(* IEC 61131-3 sources: plc-st-coding-agent/progress/evidence/f14_v14_remaining_20261113/jobs/codex_deepseek-v4pro (part 4) *)

(* ---- public-medium-04.candidate_02.st ---- *)
FUNCTION_BLOCK FB
VAR_INPUT
    TemperatureSensorInput : REAL;
    SetTemperature : REAL;
END_VAR
VAR_OUTPUT
    CurrentTemperature : REAL;
    SetTempDisplay : REAL;
    HeaterStatus : BOOL;
    OverheatProtection : BOOL;
    HeaterOutput : BOOL;
END_VAR
VAR
    tmp_SensorFault : BOOL;
    tmp_HeaterRequest : BOOL;
    tmp_OverheatLatched : BOOL;
    tmp_WasOverheat : BOOL;
    tmp_ContinuityTimer : TON;
    tmp_CoolingTimer : TON;
END_VAR

(* ENGINEERING_CONTRACT
HeaterOutput:
  ACT: TemperatureSensorInput < SetTemperature, no sensor fault, no overheat [PUB003].
  HOLD: none; recalculated each scan. OFF: equal/higher setpoint, fault, or overheat [PUB004, PUB005, PUB007].
OverheatProtection:
  ACT: heater remains on continuously for >5s, latched; HOLD: latched; OFF: auto after T#3S cooldown [PUB005].
Displays:
  CurrentTemperature mirrors sensor, SetTempDisplay mirrors setpoint, HeaterStatus mirrors HeaterOutput,
  OverheatProtection mirrors overheat latch [PUB001, PUB006].
Priority same scan: fault and overheat inhibit HeaterOutput. Sensor fault: input <0.0 or >100.0.
Units: REAL temperature values, TIME 5s/3s. Equality/manual reset unspecified; equal setpoint turns heater off.
*)
(* CONTRACT_RULES [] *)

tmp_SensorFault := (TemperatureSensorInput < 0.0) OR (TemperatureSensorInput > 100.0);
CurrentTemperature := TemperatureSensorInput;
SetTempDisplay := SetTemperature;

tmp_WasOverheat := tmp_OverheatLatched;

IF tmp_WasOverheat THEN
    tmp_CoolingTimer(IN := TRUE, PT := T#3S);
    IF tmp_CoolingTimer.Q THEN
        tmp_OverheatLatched := FALSE;
    END_IF;
END_IF;

tmp_HeaterRequest := (NOT tmp_SensorFault) AND (NOT tmp_OverheatLatched) AND (TemperatureSensorInput < SetTemperature);
HeaterOutput := tmp_HeaterRequest;

tmp_ContinuityTimer(IN := HeaterOutput, PT := T#10S);
IF tmp_ContinuityTimer.ET > T#5S THEN
    tmp_OverheatLatched := TRUE;
    HeaterOutput := FALSE;
    tmp_ContinuityTimer(IN := FALSE, PT := T#10S);
END_IF;

OverheatProtection := tmp_OverheatLatched;
HeaterStatus := HeaterOutput;

IF NOT tmp_WasOverheat THEN
    tmp_CoolingTimer(IN := tmp_OverheatLatched, PT := T#3S);
END_IF;
END_FUNCTION_BLOCK

(* ---- public-medium-04.patch_base_02.st ---- *)
FUNCTION_BLOCK FB
VAR_INPUT
    TemperatureSensorInput : REAL;
    SetTemperature : REAL;
END_VAR
VAR_OUTPUT
    CurrentTemperature : REAL;
    SetTempDisplay : REAL;
    HeaterStatus : BOOL;
    OverheatProtection : BOOL;
    HeaterOutput : BOOL;
END_VAR
VAR
    tmp_SensorFault : BOOL;
    tmp_HeaterRequest : BOOL;
    tmp_OverheatLatched : BOOL;
    tmp_WasOverheat : BOOL;
    tmp_ContinuityTimer : TON;
    tmp_CoolingTimer : TON;
END_VAR

(* ENGINEERING_CONTRACT
HeaterOutput:
  ACT: TemperatureSensorInput < SetTemperature, no sensor fault, no overheat [PUB003].
  HOLD: none; recalculated each scan. OFF: equal/higher setpoint, fault, or overheat [PUB004, PUB005, PUB007].
OverheatProtection:
  ACT: heater remains on continuously for >5s, latched; HOLD: latched; OFF: auto after T#3S cooldown [PUB005].
Displays:
  CurrentTemperature mirrors sensor, SetTempDisplay mirrors setpoint, HeaterStatus mirrors HeaterOutput,
  OverheatProtection mirrors overheat latch [PUB001, PUB006].
Priority same scan: fault and overheat inhibit HeaterOutput. Sensor fault: input <0.0 or >100.0.
Units: REAL temperature values, TIME 5s/3s. Equality/manual reset unspecified; equal setpoint turns heater off.
*)
(* CONTRACT_RULES [] *)

tmp_SensorFault := (TemperatureSensorInput < 0.0) OR (TemperatureSensorInput > 100.0);
CurrentTemperature := TemperatureSensorInput;
SetTempDisplay := SetTemperature;

tmp_WasOverheat := tmp_OverheatLatched;

IF tmp_WasOverheat THEN
    tmp_CoolingTimer(IN := TRUE, PT := T#3S);
    IF tmp_CoolingTimer.Q THEN
        tmp_OverheatLatched := FALSE;
    END_IF;
END_IF;

tmp_HeaterRequest := (NOT tmp_SensorFault) AND (NOT tmp_OverheatLatched) AND (TemperatureSensorInput < SetTemperature);
HeaterOutput := tmp_HeaterRequest;

tmp_ContinuityTimer(IN := HeaterOutput, PT := T#10S);
IF tmp_ContinuityTimer.ET > T#5S THEN
    tmp_OverheatLatched := TRUE;
    HeaterOutput := FALSE;
END_IF;

OverheatProtection := tmp_OverheatLatched;
HeaterStatus := HeaterOutput;

IF NOT tmp_WasOverheat THEN
    tmp_CoolingTimer(IN := tmp_OverheatLatched, PT := T#3S);
END_IF;
END_FUNCTION_BLOCK

(* ---- public-medium-04.raw_candidate_01.st ---- *)
FUNCTION_BLOCK FB
VAR_INPUT
    TemperatureSensorInput : REAL;
    SetTemperature : REAL;
END_VAR
VAR_OUTPUT
    CurrentTemperature : REAL;
    SetTempDisplay : REAL;
    HeaterStatus : BOOL;
    OverheatProtection : BOOL;
    HeaterOutput : BOOL;
END_VAR
VAR
    tmp_SensorFault : BOOL;
    tmp_HeaterRequest : BOOL;
    tmp_OverheatLatched : BOOL;
    tmp_WasOverheat : BOOL;
    tmp_ContinuityTimer : TON;
    tmp_CoolingTimer : TON;
END_VAR

(* ENGINEERING_CONTRACT
HeaterOutput:
  ACT: TemperatureSensorInput < SetTemperature, no sensor fault, no overheat [PUB003].
  HOLD: none; recalculated each scan. OFF: equal/higher setpoint, fault, or overheat [PUB004, PUB005, PUB007].
OverheatProtection:
  ACT: heater remains on continuously for >5s, latched; HOLD: latched; OFF: auto after T#3S cooldown [PUB005].
Displays:
  CurrentTemperature mirrors sensor, SetTempDisplay mirrors setpoint, HeaterStatus mirrors HeaterOutput,
  OverheatProtection mirrors overheat latch [PUB001, PUB006].
Priority same scan: fault and overheat inhibit HeaterOutput. Sensor fault: input <0.0 or >100.0.
Units: REAL temperature values, TIME 5s/3s. Equality/manual reset unspecified; equal setpoint turns heater off.
*)
(* CONTRACT_RULES [] *)

tmp_SensorFault := (TemperatureSensorInput < 0.0) OR (TemperatureSensorInput > 100.0);
CurrentTemperature := TemperatureSensorInput;
SetTempDisplay := SetTemperature;

tmp_WasOverheat := tmp_OverheatLatched;

IF tmp_WasOverheat THEN
    tmp_CoolingTimer(IN := TRUE, PT := T#3S);
    IF tmp_CoolingTimer.Q THEN
        tmp_OverheatLatched := FALSE;
    END_IF;
END_IF;

tmp_HeaterRequest := (NOT tmp_SensorFault) AND (NOT tmp_OverheatLatched) AND (TemperatureSensorInput < SetTemperature);
HeaterOutput := tmp_HeaterRequest;

tmp_ContinuityTimer(IN := HeaterOutput, PT := T#10S);
IF tmp_ContinuityTimer.ET > T#5S THEN
    tmp_OverheatLatched := TRUE;
    HeaterOutput := FALSE;
END_IF;

OverheatProtection := tmp_OverheatLatched;
HeaterStatus := HeaterOutput;

IF NOT tmp_WasOverheat THEN
    tmp_CoolingTimer(IN := tmp_OverheatLatched, PT := T#3S);
END_IF;
END_FUNCTION_BLOCK

(* ---- public-medium-04.raw_candidate_02.st ---- *)
FUNCTION_BLOCK FB
VAR_INPUT
    TemperatureSensorInput : REAL;
    SetTemperature : REAL;
END_VAR
VAR_OUTPUT
    CurrentTemperature : REAL;
    SetTempDisplay : REAL;
    HeaterStatus : BOOL;
    OverheatProtection : BOOL;
    HeaterOutput : BOOL;
END_VAR
VAR
    tmp_SensorFault : BOOL;
    tmp_HeaterRequest : BOOL;
    tmp_OverheatLatched : BOOL;
    tmp_WasOverheat : BOOL;
    tmp_ContinuityTimer : TON;
    tmp_CoolingTimer : TON;
END_VAR

(* ENGINEERING_CONTRACT
HeaterOutput:
  ACT: TemperatureSensorInput < SetTemperature, no sensor fault, no overheat [PUB003].
  HOLD: none; recalculated each scan. OFF: equal/higher setpoint, fault, or overheat [PUB004, PUB005, PUB007].
OverheatProtection:
  ACT: heater remains on continuously for >5s, latched; HOLD: latched; OFF: auto after T#3S cooldown [PUB005].
Displays:
  CurrentTemperature mirrors sensor, SetTempDisplay mirrors setpoint, HeaterStatus mirrors HeaterOutput,
  OverheatProtection mirrors overheat latch [PUB001, PUB006].
Priority same scan: fault and overheat inhibit HeaterOutput. Sensor fault: input <0.0 or >100.0.
Units: REAL temperature values, TIME 5s/3s. Equality/manual reset unspecified; equal setpoint turns heater off.
*)
(* CONTRACT_RULES [] *)

tmp_SensorFault := (TemperatureSensorInput < 0.0) OR (TemperatureSensorInput > 100.0);
CurrentTemperature := TemperatureSensorInput;
SetTempDisplay := SetTemperature;

tmp_WasOverheat := tmp_OverheatLatched;

IF tmp_WasOverheat THEN
    tmp_CoolingTimer(IN := TRUE, PT := T#3S);
    IF tmp_CoolingTimer.Q THEN
        tmp_OverheatLatched := FALSE;
    END_IF;
END_IF;

tmp_HeaterRequest := (NOT tmp_SensorFault) AND (NOT tmp_OverheatLatched) AND (TemperatureSensorInput < SetTemperature);
HeaterOutput := tmp_HeaterRequest;

tmp_ContinuityTimer(IN := HeaterOutput, PT := T#10S);
IF tmp_ContinuityTimer.ET > T#5S THEN
    tmp_OverheatLatched := TRUE;
    HeaterOutput := FALSE;
    tmp_ContinuityTimer(IN := FALSE, PT := T#10S);
END_IF;

OverheatProtection := tmp_OverheatLatched;
HeaterStatus := HeaterOutput;

IF NOT tmp_WasOverheat THEN
    tmp_CoolingTimer(IN := tmp_OverheatLatched, PT := T#3S);
END_IF;
END_FUNCTION_BLOCK

(* ---- public-medium-05.candidate_01.st ---- *)
TYPE LineTarget : (TargetNone, TargetB, TargetC);
END_TYPE;

FUNCTION_BLOCK ProductionLineControl
VAR_INPUT
    Mode : BOOL;
    ForwardButton : BOOL;
    ReverseButton : BOOL;
    SensorA : BOOL;
    SensorB : BOOL;
    SensorC : BOOL;
    ButtonA : BOOL;
    ButtonB : BOOL;
    ButtonC : BOOL;
END_VAR
VAR_OUTPUT
    MotorForward : BOOL;
    MotorReverse : BOOL;
    CompletionLight : BOOL;
END_VAR
VAR
    local_target : LineTarget := TargetNone;
    completionLatched : BOOL := FALSE;
END_VAR

(* ENGINEERING_CONTRACT
MotorForward auto: activated by ButtonA at SensorA or ButtonB at SensorB; held until target SensorB/C.
MotorForward manual: follows ForwardButton while ReverseButton is FALSE; both conflict outputs inhibited.
MotorReverse manual: follows ReverseButton while ForwardButton is FALSE; auto mode holds MotorReverse OFF.
CompletionLight: latched TRUE on Mode & SensorC & ButtonC; retained until SensorC becomes FALSE.
Same-scan priority: SensorC, then SensorB, then SensorA; arrival plus next button uses final current inputs.
Mode-transition retention is unspecified; auto target and completion state are retained when mode changes.
Units/boundaries: BOOL logic only; no time or arithmetic boundaries.
*)

(* CONTRACT_RULES [] *)

IF Mode THEN
    CASE local_target OF
        TargetNone:
            IF SensorC THEN
                IF ButtonC THEN
                    completionLatched := TRUE;
                END_IF;
            ELSIF SensorB THEN
                IF ButtonB THEN
                    local_target := TargetC;
                END_IF;
            ELSIF SensorA AND ButtonA THEN
                local_target := TargetB;
            END_IF;

        TargetB:
            IF SensorC THEN
                local_target := TargetNone;
                IF ButtonC THEN
                    completionLatched := TRUE;
                END_IF;
            ELSIF SensorB THEN
                local_target := TargetNone;
                IF ButtonB THEN
                    local_target := TargetC;
                END_IF;
            END_IF;

        TargetC:
            IF SensorC THEN
                local_target := TargetNone;
                IF ButtonC THEN
                    completionLatched := TRUE;
                END_IF;
            END_IF;
    END_CASE;

    IF local_target <> TargetNone THEN
        MotorForward := TRUE;
    ELSE
        MotorForward := FALSE;
    END_IF;
    MotorReverse := FALSE;
ELSE
    MotorForward := ForwardButton AND NOT ReverseButton;
    MotorReverse := ReverseButton AND NOT ForwardButton;
END_IF;

IF NOT SensorC THEN
    completionLatched := FALSE;
END_IF;

CompletionLight := completionLatched;

END_FUNCTION_BLOCK

(* ---- public-medium-05.raw_candidate_01.st ---- *)
TYPE LineTarget : (TargetNone, TargetB, TargetC);
END_TYPE

FUNCTION_BLOCK ProductionLineControl
VAR_INPUT
    Mode : BOOL;
    ForwardButton : BOOL;
    ReverseButton : BOOL;
    SensorA : BOOL;
    SensorB : BOOL;
    SensorC : BOOL;
    ButtonA : BOOL;
    ButtonB : BOOL;
    ButtonC : BOOL;
END_VAR
VAR_OUTPUT
    MotorForward : BOOL;
    MotorReverse : BOOL;
    CompletionLight : BOOL;
END_VAR
VAR
    local_target : LineTarget := TargetNone;
    completionLatched : BOOL := FALSE;
END_VAR

(* ENGINEERING_CONTRACT
MotorForward auto: activated by ButtonA at SensorA or ButtonB at SensorB; held until target SensorB/C.
MotorForward manual: follows ForwardButton while ReverseButton is FALSE; both conflict outputs inhibited.
MotorReverse manual: follows ReverseButton while ForwardButton is FALSE; auto mode holds MotorReverse OFF.
CompletionLight: latched TRUE on Mode & SensorC & ButtonC; retained until SensorC becomes FALSE.
Same-scan priority: SensorC, then SensorB, then SensorA; arrival plus next button uses final current inputs.
Mode-transition retention is unspecified; auto target and completion state are retained when mode changes.
Units/boundaries: BOOL logic only; no time or arithmetic boundaries.
*)

(* CONTRACT_RULES [] *)

IF Mode THEN
    CASE local_target OF
        TargetNone:
            IF SensorC THEN
                IF ButtonC THEN
                    completionLatched := TRUE;
                END_IF;
            ELSIF SensorB THEN
                IF ButtonB THEN
                    local_target := TargetC;
                END_IF;
            ELSIF SensorA AND ButtonA THEN
                local_target := TargetB;
            END_IF;

        TargetB:
            IF SensorC THEN
                local_target := TargetNone;
                IF ButtonC THEN
                    completionLatched := TRUE;
                END_IF;
            ELSIF SensorB THEN
                local_target := TargetNone;
                IF ButtonB THEN
                    local_target := TargetC;
                END_IF;
            END_IF;

        TargetC:
            IF SensorC THEN
                local_target := TargetNone;
                IF ButtonC THEN
                    completionLatched := TRUE;
                END_IF;
            END_IF;
    END_CASE;

    IF local_target <> TargetNone THEN
        MotorForward := TRUE;
    ELSE
        MotorForward := FALSE;
    END_IF;
    MotorReverse := FALSE;
ELSE
    MotorForward := ForwardButton AND NOT ReverseButton;
    MotorReverse := ReverseButton AND NOT ForwardButton;
END_IF;

IF NOT SensorC THEN
    completionLatched := FALSE;
END_IF;

CompletionLight := completionLatched;

END_FUNCTION_BLOCK

(* ---- public-medium-06.candidate_01.st ---- *)
FUNCTION_BLOCK FB_SlabThicknessAlarmHistory
(* ENGINEERING_CONTRACT
THICKNESS_ALARM: set on valid-fault rising edge; TON holds >=500 ms; current fault keeps it on; signal invalid clears (PUB001,PUB004).
Slab_Fault_Counter: increments once per valid-fault rising edge; retained otherwise; UINT wrap unspecified (PUB002).
Slab_Fault_History: newest stored at index 0, older entries shifted upward, five entries retained; zero at power-up (PUB002,PUB005).
Slab_Runtime_Accumulator: adds TIME_TO_LTIME(CycleTime) only when CUTTING_RUN AND valid AND NOT fault; retained otherwise (PUB003).
Invalid/power-up: alarm false and timer cleared; no record or runtime accumulation while signal invalid (PUB004,PUB005).
Same-scan priority: record/alarm edge processed before runtime condition, so a faulted scan adds no normal runtime.
Hold timer: retriggerable; edge reset precedes enabled TON call; Q completion releases hold on the following valid scan.
Units/boundaries: hold threshold T#500MS inclusive via TON >=; runtime LTIME nanoseconds; history index 0 newest.
*)
(* CONTRACT_RULES [] *)
VAR_INPUT
    THICKNESS_FAULT : BOOL;
    THICKNESS_SIGNAL_VALID : BOOL;
    CUTTING_RUN : BOOL;
    FaultTimestamp : DINT;
    CycleTime : TIME;
END_VAR
VAR_OUTPUT
    THICKNESS_ALARM : BOOL;
    Slab_Fault_Counter : UINT;
    Slab_Runtime_Accumulator : LTIME;
    Slab_Fault_History : ARRAY[0..4] OF DINT;
END_VAR
VAR
    local_valid_fault : BOOL;
    local_fault_rise : R_TRIG;
    local_alarm_timer : TON;
    local_hold_active : BOOL;
    local_cycle_ltime : LTIME;
    local_i : INT;
END_VAR

local_valid_fault := THICKNESS_SIGNAL_VALID AND THICKNESS_FAULT;
local_fault_rise(CLK := local_valid_fault);
local_cycle_ltime := TIME_TO_LTIME(CycleTime);

IF NOT THICKNESS_SIGNAL_VALID THEN
    THICKNESS_ALARM := FALSE;
    local_hold_active := FALSE;
    local_alarm_timer(IN := FALSE, PT := T#500MS);
ELSIF local_fault_rise.Q THEN
    Slab_Fault_Counter := Slab_Fault_Counter + UINT#1;

    FOR local_i := 4 TO 1 BY -1 DO
        Slab_Fault_History[local_i] := Slab_Fault_History[local_i - 1];
    END_FOR;

    Slab_Fault_History[0] := FaultTimestamp;
    local_hold_active := TRUE;
    local_alarm_timer(IN := FALSE, PT := T#500MS);
END_IF;

IF THICKNESS_SIGNAL_VALID THEN
    IF local_alarm_timer.Q THEN
        local_hold_active := FALSE;
    END_IF;

    local_alarm_timer(IN := local_hold_active, PT := T#500MS);

    THICKNESS_ALARM := THICKNESS_FAULT OR local_hold_active;
END_IF;

IF CUTTING_RUN AND THICKNESS_SIGNAL_VALID AND NOT THICKNESS_FAULT THEN
    Slab_Runtime_Accumulator := Slab_Runtime_Accumulator + local_cycle_ltime;
END_IF;

END_FUNCTION_BLOCK

(* ---- public-medium-06.raw_candidate_01.st ---- *)
FUNCTION_BLOCK FB_SlabThicknessAlarmHistory
(* ENGINEERING_CONTRACT
THICKNESS_ALARM: set on valid-fault rising edge; TON holds >=500 ms; current fault keeps it on; signal invalid clears (PUB001,PUB004).
Slab_Fault_Counter: increments once per valid-fault rising edge; retained otherwise; UINT wrap unspecified (PUB002).
Slab_Fault_History: newest stored at index 0, older entries shifted upward, five entries retained; zero at power-up (PUB002,PUB005).
Slab_Runtime_Accumulator: adds TIME_TO_LTIME(CycleTime) only when CUTTING_RUN AND valid AND NOT fault; retained otherwise (PUB003).
Invalid/power-up: alarm false and timer cleared; no record or runtime accumulation while signal invalid (PUB004,PUB005).
Same-scan priority: record/alarm edge processed before runtime condition, so a faulted scan adds no normal runtime.
Hold timer: retriggerable; edge reset precedes enabled TON call; Q completion releases hold on the following valid scan.
Units/boundaries: hold threshold T#500MS inclusive via TON >=; runtime LTIME nanoseconds; history index 0 newest.
*)
(* CONTRACT_RULES [] *)
VAR_INPUT
    THICKNESS_FAULT : BOOL;
    THICKNESS_SIGNAL_VALID : BOOL;
    CUTTING_RUN : BOOL;
    FaultTimestamp : DINT;
    CycleTime : TIME;
END_VAR
VAR_OUTPUT
    THICKNESS_ALARM : BOOL;
    Slab_Fault_Counter : UINT;
    Slab_Runtime_Accumulator : LTIME;
    Slab_Fault_History : ARRAY[0..4] OF DINT;
END_VAR
VAR
    local_valid_fault : BOOL;
    local_fault_rise : R_TRIG;
    local_alarm_timer : TON;
    local_hold_active : BOOL;
    local_cycle_ltime : LTIME;
    local_i : INT;
END_VAR

local_valid_fault := THICKNESS_SIGNAL_VALID AND THICKNESS_FAULT;
local_fault_rise(CLK := local_valid_fault);
local_cycle_ltime := TIME_TO_LTIME(CycleTime);

IF NOT THICKNESS_SIGNAL_VALID THEN
    THICKNESS_ALARM := FALSE;
    local_hold_active := FALSE;
    local_alarm_timer(IN := FALSE, PT := T#500MS);
ELSIF local_fault_rise.Q THEN
    Slab_Fault_Counter := Slab_Fault_Counter + UINT#1;

    FOR local_i := 4 TO 1 BY -1 DO
        Slab_Fault_History[local_i] := Slab_Fault_History[local_i - 1];
    END_FOR;

    Slab_Fault_History[0] := FaultTimestamp;
    local_hold_active := TRUE;
    local_alarm_timer(IN := FALSE, PT := T#500MS);
END_IF;

IF THICKNESS_SIGNAL_VALID THEN
    IF local_alarm_timer.Q THEN
        local_hold_active := FALSE;
    END_IF;

    local_alarm_timer(IN := local_hold_active, PT := T#500MS);

    THICKNESS_ALARM := THICKNESS_FAULT OR local_hold_active;
END_IF;

IF CUTTING_RUN AND THICKNESS_SIGNAL_VALID AND NOT THICKNESS_FAULT THEN
    Slab_Runtime_Accumulator := Slab_Runtime_Accumulator + local_cycle_ltime;
END_IF;

END_FUNCTION_BLOCK

(* ---- public-medium-07.candidate_01.st ---- *)
FUNCTION_BLOCK HVACMultiModeControl
VAR_INPUT
    OCCUPANCY_DETECTED : BOOL;
    ENERGY_SAVING_MODE : BOOL;
    HVAC_MODE_SELECTOR : INT;
END_VAR
VAR_OUTPUT
    SUPPLY_FAN_RUN : BOOL;
    TEMP_SETPOINT_ADJUST : INT;
END_VAR
VAR
    tmp_Delay : TON;
    tmp_Enable : BOOL;
    tmp_Adjust : INT;
END_VAR

(* ENGINEERING_CONTRACT
   SUPPLY_FAN_RUN [PUB002, PUB005]: enabled only while occupancy exists
   and HVAC_MODE_SELECTOR <> 3; TON 30 s drives the output. Losing the
   enable condition stops output and resets timing on the same scan;
   recovery requires a complete new 30 s interval.
   TEMP_SETPOINT_ADJUST [PUB003, PUB004]: recomputed each scan. Auto is
   0/3/2, Comfort 0/1, Economy 0/4, Night 4; energy saving affects Auto
   only. Result is clamped to [-4, +4] °C.
   Init state: outputs OFF and 0 at power-up; invalid selector uses 0 °C.
*)

(* CONTRACT_RULES [] *)

SUPPLY_FAN_RUN := FALSE;
TEMP_SETPOINT_ADJUST := 0;

tmp_Enable := OCCUPANCY_DETECTED AND (HVAC_MODE_SELECTOR <> 3);
tmp_Delay(IN := tmp_Enable, PT := T#30S);
SUPPLY_FAN_RUN := tmp_Delay.Q;

CASE HVAC_MODE_SELECTOR OF
    0:
        IF OCCUPANCY_DETECTED THEN
            tmp_Adjust := 0;
        ELSIF ENERGY_SAVING_MODE THEN
            tmp_Adjust := 3;
        ELSE
            tmp_Adjust := 2;
        END_IF;
    1:
        IF OCCUPANCY_DETECTED THEN
            tmp_Adjust := 0;
        ELSE
            tmp_Adjust := 1;
        END_IF;
    2:
        IF OCCUPANCY_DETECTED THEN
            tmp_Adjust := 0;
        ELSE
            tmp_Adjust := 4;
        END_IF;
    3:
        tmp_Adjust := 4;
    ELSE
        tmp_Adjust := 0;
END_CASE;

IF tmp_Adjust < -4 THEN
    tmp_Adjust := -4;
ELSIF tmp_Adjust > 4 THEN
    tmp_Adjust := 4;
END_IF;

TEMP_SETPOINT_ADJUST := tmp_Adjust;
END_FUNCTION_BLOCK

(* ---- public-medium-07.raw_candidate_01.st ---- *)
FUNCTION_BLOCK HVACMultiModeControl
VAR_INPUT
    OCCUPANCY_DETECTED : BOOL;
    ENERGY_SAVING_MODE : BOOL;
    HVAC_MODE_SELECTOR : INT;
END_VAR
VAR_OUTPUT
    SUPPLY_FAN_RUN : BOOL;
    TEMP_SETPOINT_ADJUST : INT;
END_VAR
VAR
    tmp_Delay : TON;
    tmp_Enable : BOOL;
    tmp_Adjust : INT;
END_VAR

(* ENGINEERING_CONTRACT
   SUPPLY_FAN_RUN [PUB002, PUB005]: enabled only while occupancy exists
   and HVAC_MODE_SELECTOR <> 3; TON 30 s drives the output. Losing the
   enable condition stops output and resets timing on the same scan;
   recovery requires a complete new 30 s interval.
   TEMP_SETPOINT_ADJUST [PUB003, PUB004]: recomputed each scan. Auto is
   0/3/2, Comfort 0/1, Economy 0/4, Night 4; energy saving affects Auto
   only. Result is clamped to [-4, +4] °C.
   Init state: outputs OFF and 0 at power-up; invalid selector uses 0 °C.
*)

(* CONTRACT_RULES [] *)

SUPPLY_FAN_RUN := FALSE;
TEMP_SETPOINT_ADJUST := 0;

tmp_Enable := OCCUPANCY_DETECTED AND (HVAC_MODE_SELECTOR <> 3);
tmp_Delay(IN := tmp_Enable, PT := T#30S);
SUPPLY_FAN_RUN := tmp_Delay.Q;

CASE HVAC_MODE_SELECTOR OF
    0:
        IF OCCUPANCY_DETECTED THEN
            tmp_Adjust := 0;
        ELSIF ENERGY_SAVING_MODE THEN
            tmp_Adjust := 3;
        ELSE
            tmp_Adjust := 2;
        END_IF;
    1:
        IF OCCUPANCY_DETECTED THEN
            tmp_Adjust := 0;
        ELSE
            tmp_Adjust := 1;
        END_IF;
    2:
        IF OCCUPANCY_DETECTED THEN
            tmp_Adjust := 0;
        ELSE
            tmp_Adjust := 4;
        END_IF;
    3:
        tmp_Adjust := 4;
    ELSE
        tmp_Adjust := 0;
END_CASE;

IF tmp_Adjust < -4 THEN
    tmp_Adjust := -4;
ELSIF tmp_Adjust > 4 THEN
    tmp_Adjust := 4;
END_IF;

TEMP_SETPOINT_ADJUST := tmp_Adjust;
END_FUNCTION_BLOCK

(* ---- public-medium-08.candidate_01.st ---- *)
(* ENGINEERING_CONTRACT
ipValue is combinational and recomputed every scan; no retention (PUB003).
Activation: exactly three periods and four nonempty all-digit segments (PUB001/PUB002).
Invalid/reset: len<7, len>15, nondigit, extra/missing dot, empty segment, or value>255 => 0 (PUB001/PUB003/PUB004).
Assemble seg1<<24 | seg2<<16 | seg3<<8 | seg4 (PUB002/PUB004).
0.0.0.0 and invalid both produce 0, distinguished only by structural checks.
Malformed condition dominates valid assembly; final ipValue is 0.
Unspecified: leading zeros are accepted; whitespace/sign characters are rejected.
*)
(* CONTRACT_RULES [] *)
FUNCTION_BLOCK FB_IPv4Parser
VAR_INPUT
    ipText : STRING(254);
END_VAR
VAR_OUTPUT
    ipValue : UDINT;
END_VAR
VAR
    tmp_len : INT;
    tmp_idx : INT;
    tmp_char : BYTE;
    tmp_digit : UDINT;
    tmp_seg_value : UDINT;
    tmp_new_value : UDINT;
    tmp_addr : UDINT;
    tmp_seg_count : INT;
    tmp_in_segment : BOOL;
    tmp_valid : BOOL;
END_VAR

tmp_len := LEN(ipText);
tmp_valid := (tmp_len >= 7) AND (tmp_len <= 15);
tmp_addr := UDINT#0;
tmp_seg_count := 0;
tmp_in_segment := FALSE;
tmp_seg_value := UDINT#0;
tmp_new_value := UDINT#0;

IF tmp_valid THEN
    FOR tmp_idx := 0 TO tmp_len - 1 DO
        tmp_char := ipText[tmp_idx];

        IF (tmp_char >= 48) AND (tmp_char <= 57) THEN
            tmp_in_segment := TRUE;
            IF tmp_seg_value <= UDINT#255 THEN
                tmp_digit := BYTE_TO_UDINT(tmp_char) - UDINT#48;
                tmp_new_value := (tmp_seg_value * UDINT#10) + tmp_digit;
                IF tmp_new_value > UDINT#255 THEN
                    tmp_seg_value := UDINT#256;
                    tmp_valid := FALSE;
                ELSE
                    tmp_seg_value := tmp_new_value;
                END_IF;
            END_IF;
        ELSIF tmp_char = 46 THEN
            IF tmp_in_segment THEN
                tmp_seg_count := tmp_seg_count + 1;
                IF tmp_seg_count > 3 THEN
                    tmp_valid := FALSE;
                END_IF;
                tmp_addr := SHL(tmp_addr, 8) OR tmp_seg_value;
                tmp_seg_value := UDINT#0;
                tmp_in_segment := FALSE;
            ELSE
                tmp_valid := FALSE;
            END_IF;
        ELSE
            tmp_valid := FALSE;
        END_IF;
    END_FOR;

    IF tmp_in_segment THEN
        tmp_addr := SHL(tmp_addr, 8) OR tmp_seg_value;
        tmp_seg_count := tmp_seg_count + 1;
        tmp_in_segment := FALSE;
    ELSE
        tmp_valid := FALSE;
    END_IF;
END_IF;

IF tmp_valid AND (tmp_seg_count = 4) THEN
    ipValue := tmp_addr;
ELSE
    ipValue := UDINT#0;
END_IF;

END_FUNCTION_BLOCK

(* ---- public-medium-08.raw_candidate_01.st ---- *)
(* ENGINEERING_CONTRACT
ipValue is combinational and recomputed every scan; no retention (PUB003).
Activation: exactly three periods and four nonempty all-digit segments (PUB001/PUB002).
Invalid/reset: len<7, len>15, nondigit, extra/missing dot, empty segment, or value>255 => 0 (PUB001/PUB003/PUB004).
Assemble seg1<<24 | seg2<<16 | seg3<<8 | seg4 (PUB002/PUB004).
0.0.0.0 and invalid both produce 0, distinguished only by structural checks.
Malformed condition dominates valid assembly; final ipValue is 0.
Unspecified: leading zeros are accepted; whitespace/sign characters are rejected.
*)
(* CONTRACT_RULES [] *)
FUNCTION_BLOCK FB_IPv4Parser
VAR_INPUT
    ipText : STRING(254);
END_VAR
VAR_OUTPUT
    ipValue : UDINT;
END_VAR
VAR
    tmp_len : INT;
    tmp_idx : INT;
    tmp_char : BYTE;
    tmp_digit : UDINT;
    tmp_seg_value : UDINT;
    tmp_new_value : UDINT;
    tmp_addr : UDINT;
    tmp_seg_count : INT;
    tmp_in_segment : BOOL;
    tmp_valid : BOOL;
END_VAR

tmp_len := LEN(ipText);
tmp_valid := (tmp_len >= 7) AND (tmp_len <= 15);
tmp_addr := UDINT#0;
tmp_seg_count := 0;
tmp_in_segment := FALSE;
tmp_seg_value := UDINT#0;
tmp_new_value := UDINT#0;

IF tmp_valid THEN
    FOR tmp_idx := 0 TO tmp_len - 1 DO
        tmp_char := ipText[tmp_idx];

        IF (tmp_char >= 48) AND (tmp_char <= 57) THEN
            tmp_in_segment := TRUE;
            IF tmp_seg_value <= UDINT#255 THEN
                tmp_digit := BYTE_TO_UDINT(tmp_char) - UDINT#48;
                tmp_new_value := (tmp_seg_value * UDINT#10) + tmp_digit;
                IF tmp_new_value > UDINT#255 THEN
                    tmp_seg_value := UDINT#256;
                    tmp_valid := FALSE;
                ELSE
                    tmp_seg_value := tmp_new_value;
                END_IF;
            END_IF;
        ELSIF tmp_char = 46 THEN
            IF tmp_in_segment THEN
                tmp_seg_count := tmp_seg_count + 1;
                IF tmp_seg_count > 3 THEN
                    tmp_valid := FALSE;
                END_IF;
                tmp_addr := SHL(tmp_addr, 8) OR tmp_seg_value;
                tmp_seg_value := UDINT#0;
                tmp_in_segment := FALSE;
            ELSE
                tmp_valid := FALSE;
            END_IF;
        ELSE
            tmp_valid := FALSE;
        END_IF;
    END_FOR;

    IF tmp_in_segment THEN
        tmp_addr := SHL(tmp_addr, 8) OR tmp_seg_value;
        tmp_seg_count := tmp_seg_count + 1;
        tmp_in_segment := FALSE;
    ELSE
        tmp_valid := FALSE;
    END_IF;
END_IF;

IF tmp_valid AND (tmp_seg_count = 4) THEN
    ipValue := tmp_addr;
ELSE
    ipValue := UDINT#0;
END_IF;

END_FUNCTION_BLOCK

(* ---- self-easy-01.candidate_01.st ---- *)
FUNCTION_BLOCK FB
(* ENGINEERING_CONTRACT
   avgOut is a retained process value written only on an active valid average scan.
   Activation: enable AND avgEnable AND count >= 1.
   Hold: avgOut remains unchanged when enable=FALSE, avgEnable=FALSE, or count<=0.
   Explicit reset: none specified.
   Same-scan priority: active valid calculation wins; invalid/disabled leaves avgOut unchanged.
   Boundaries: count<1 means no update; count in 1..8 uses count samples; count>8 clips to 8.
   Units: INT samples summed in DINT, divided in REAL; boundary time/scan: current cycle.
   Cite: PUB001-PUB027 behavior clauses; formal S1-S6.
*)
(* CONTRACT_RULES [] *)
VAR_INPUT
    enable : BOOL;
    values : ARRAY[1..8] OF INT;
    count : INT;
    avgEnable : BOOL;
END_VAR
VAR_OUTPUT
    avgOut : REAL;
END_VAR
VAR
    tmp_sum : DINT;
    tmp_count : INT;
    tmp_i : INT;
END_VAR

IF enable AND avgEnable AND (count >= 1) THEN
    tmp_count := count;
    IF tmp_count > 8 THEN
        tmp_count := 8;
    END_IF;

    tmp_sum := 0;
    FOR tmp_i := 1 TO tmp_count DO
        tmp_sum := tmp_sum + INT_TO_DINT(values[tmp_i]);
    END_FOR;

    avgOut := DINT_TO_REAL(tmp_sum) / INT_TO_REAL(tmp_count);
END_IF;

END_FUNCTION_BLOCK

(* ---- self-easy-01.raw_candidate_01.st ---- *)
FUNCTION_BLOCK FB
(* ENGINEERING_CONTRACT
   avgOut is a retained process value written only on an active valid average scan.
   Activation: enable AND avgEnable AND count >= 1.
   Hold: avgOut remains unchanged when enable=FALSE, avgEnable=FALSE, or count<=0.
   Explicit reset: none specified.
   Same-scan priority: active valid calculation wins; invalid/disabled leaves avgOut unchanged.
   Boundaries: count<1 means no update; count in 1..8 uses count samples; count>8 clips to 8.
   Units: INT samples summed in DINT, divided in REAL; boundary time/scan: current cycle.
   Cite: PUB001-PUB027 behavior clauses; formal S1-S6.
*)
(* CONTRACT_RULES [] *)
VAR_INPUT
    enable : BOOL;
    values : ARRAY[1..8] OF INT;
    count : INT;
    avgEnable : BOOL;
END_VAR
VAR_OUTPUT
    avgOut : REAL;
END_VAR
VAR
    tmp_sum : DINT;
    tmp_count : INT;
    tmp_i : INT;
END_VAR

IF enable AND avgEnable AND (count >= 1) THEN
    tmp_count := count;
    IF tmp_count > 8 THEN
        tmp_count := 8;
    END_IF;

    tmp_sum := 0;
    FOR tmp_i := 1 TO tmp_count DO
        tmp_sum := tmp_sum + INT_TO_DINT(values[tmp_i]);
    END_FOR;

    avgOut := DINT_TO_REAL(tmp_sum) / INT_TO_REAL(tmp_count);
END_IF;

END_FUNCTION_BLOCK

(* ---- self-easy-02.candidate_01.st ---- *)
FUNCTION_BLOCK FB

(* ENGINEERING_CONTRACT
   alarms: latch immediately on their own danger condition, retain until a new
           resetBtn rising edge occurs while the condition is gone; dangerous
           condition has priority on the same scan.
   reset edge: detected from resetBtn TRUE and previous scan resetBtn FALSE;
                prevResetBtn is updated at the end of every scan.
   pumpRun: combinational after alarm update; TRUE iff inletPermit AND no alarm.
   outletValveOpen: combinational; TRUE iff low alarm is FALSE.
   tankLevel units: percent; thresholds are >= 85.0 for high and <= 15.0 for low.
   outletFlow: observed only, does not affect outputs.
*)

VAR_INPUT
    tankLevel : REAL;    (* 0..100 % *)
    outletFlow : REAL;   (* m3/h, reserved observation input *)
    inletPermit : BOOL;
    resetBtn : BOOL;
END_VAR

VAR_OUTPUT
    pumpRun : BOOL;
    alarmHigh : BOOL;
    alarmLow : BOOL;
    outletValveOpen : BOOL;
END_VAR

VAR
    local_prevResetBtn : BOOL := FALSE;
    local_risingReset : BOOL;
    tmp_highState : BOOL := FALSE;
    tmp_lowState : BOOL := FALSE;
END_VAR

(* CONTRACT_RULES [] *)

local_risingReset := resetBtn AND NOT local_prevResetBtn;

(* High alarm: danger condition sets and latches. *)
IF tankLevel >= 85.0 THEN
    tmp_highState := TRUE;
ELSIF local_risingReset THEN
    tmp_highState := FALSE;
END_IF;

(* Low alarm: danger condition sets and latches. *)
IF tankLevel <= 15.0 THEN
    tmp_lowState := TRUE;
ELSIF local_risingReset THEN
    tmp_lowState := FALSE;
END_IF;

alarmHigh := tmp_highState;
alarmLow := tmp_lowState;

pumpRun := inletPermit AND NOT alarmHigh AND NOT alarmLow;
outletValveOpen := NOT alarmLow;

local_prevResetBtn := resetBtn;

END_FUNCTION_BLOCK

(* ---- self-easy-02.raw_candidate_01.st ---- *)
FUNCTION_BLOCK FB

(* ENGINEERING_CONTRACT
   alarms: latch immediately on their own danger condition, retain until a new
           resetBtn rising edge occurs while the condition is gone; dangerous
           condition has priority on the same scan.
   reset edge: detected from resetBtn TRUE and previous scan resetBtn FALSE;
                prevResetBtn is updated at the end of every scan.
   pumpRun: combinational after alarm update; TRUE iff inletPermit AND no alarm.
   outletValveOpen: combinational; TRUE iff low alarm is FALSE.
   tankLevel units: percent; thresholds are >= 85.0 for high and <= 15.0 for low.
   outletFlow: observed only, does not affect outputs.
*)

VAR_INPUT
    tankLevel : REAL;    (* 0..100 % *)
    outletFlow : REAL;   (* m3/h, reserved observation input *)
    inletPermit : BOOL;
    resetBtn : BOOL;
END_VAR

VAR_OUTPUT
    pumpRun : BOOL;
    alarmHigh : BOOL;
    alarmLow : BOOL;
    outletValveOpen : BOOL;
END_VAR

VAR
    local_prevResetBtn : BOOL := FALSE;
    local_risingReset : BOOL;
    tmp_highState : BOOL := FALSE;
    tmp_lowState : BOOL := FALSE;
END_VAR

(* CONTRACT_RULES [] *)

local_risingReset := resetBtn AND NOT local_prevResetBtn;

(* High alarm: danger condition sets and latches. *)
IF tankLevel >= 85.0 THEN
    tmp_highState := TRUE;
ELSIF local_risingReset THEN
    tmp_highState := FALSE;
END_IF;

(* Low alarm: danger condition sets and latches. *)
IF tankLevel <= 15.0 THEN
    tmp_lowState := TRUE;
ELSIF local_risingReset THEN
    tmp_lowState := FALSE;
END_IF;

alarmHigh := tmp_highState;
alarmLow := tmp_lowState;

pumpRun := inletPermit AND NOT alarmHigh AND NOT alarmLow;
outletValveOpen := NOT alarmLow;

local_prevResetBtn := resetBtn;

END_FUNCTION_BLOCK

(* ---- self-hard-01.candidate_01.st ---- *)
(*
ENGINEERING_CONTRACT
 alarmActive: set=flowLow (PUB005); hold while unacknowledged despite flow loss (PUB006);
 clear=rising ack with flowLow=FALSE, or condition loss after confirmed-active state (PUB007/S6);
 evaluates current flowLow and rising ack in the same scan.
 alarmAcked: set=flow loss while active-unacknowledged (PUB006), rising ack with flowLow (PUB007),
 or sustained confirmation (LTL S7); clear when alarmActive becomes FALSE.
 highHigh: set/reset=!sensorOK in the same scan (PUB008-PUB009); independent of low outputs.
 Priority/units: highHigh and low-alarm outputs may be TRUE simultaneously; BOOL states; one-scan ack edge.
*)
(* CONTRACT_RULES [] *)
FUNCTION_BLOCK FB
VAR_INPUT
    flowLow : BOOL;
    ackBtn : BOOL;
    sensorOK : BOOL;
END_VAR
VAR_OUTPUT
    alarmActive : BOOL;
    alarmAcked : BOOL;
    highHigh : BOOL;
END_VAR
VAR
    local_PrevAckBtn : BOOL := FALSE;
    local_PrevFlowLow : BOOL := FALSE;
    local_PrevAlarmActive : BOOL := FALSE;
    local_PrevAlarmAcked : BOOL := FALSE;
    local_RisingAckBtn : BOOL := FALSE;
END_VAR

local_RisingAckBtn := ackBtn AND NOT local_PrevAckBtn;

alarmActive := flowLow OR
               (local_PrevAlarmActive AND
                NOT local_RisingAckBtn AND
                NOT (local_PrevFlowLow AND local_PrevAlarmAcked));

alarmAcked := alarmActive AND
              (NOT flowLow OR
               local_RisingAckBtn OR
               (local_PrevFlowLow AND local_PrevAlarmActive AND local_PrevAlarmAcked));

highHigh := NOT sensorOK;

local_PrevAckBtn := ackBtn;
local_PrevFlowLow := flowLow;
local_PrevAlarmActive := alarmActive;
local_PrevAlarmAcked := alarmAcked;

END_FUNCTION_BLOCK

(* ---- self-hard-01.raw_candidate_01.st ---- *)
(*
ENGINEERING_CONTRACT
 alarmActive: set=flowLow (PUB005); hold while unacknowledged despite flow loss (PUB006);
 clear=rising ack with flowLow=FALSE, or condition loss after confirmed-active state (PUB007/S6);
 evaluates current flowLow and rising ack in the same scan.
 alarmAcked: set=flow loss while active-unacknowledged (PUB006), rising ack with flowLow (PUB007),
 or sustained confirmation (LTL S7); clear when alarmActive becomes FALSE.
 highHigh: set/reset=!sensorOK in the same scan (PUB008-PUB009); independent of low outputs.
 Priority/units: highHigh and low-alarm outputs may be TRUE simultaneously; BOOL states; one-scan ack edge.
*)
(* CONTRACT_RULES [] *)
FUNCTION_BLOCK FB
VAR_INPUT
    flowLow : BOOL;
    ackBtn : BOOL;
    sensorOK : BOOL;
END_VAR
VAR_OUTPUT
    alarmActive : BOOL;
    alarmAcked : BOOL;
    highHigh : BOOL;
END_VAR
VAR
    local_PrevAckBtn : BOOL := FALSE;
    local_PrevFlowLow : BOOL := FALSE;
    local_PrevAlarmActive : BOOL := FALSE;
    local_PrevAlarmAcked : BOOL := FALSE;
    local_RisingAckBtn : BOOL := FALSE;
END_VAR

local_RisingAckBtn := ackBtn AND NOT local_PrevAckBtn;

alarmActive := flowLow OR
               (local_PrevAlarmActive AND
                NOT local_RisingAckBtn AND
                NOT (local_PrevFlowLow AND local_PrevAlarmAcked));

alarmAcked := alarmActive AND
              (NOT flowLow OR
               local_RisingAckBtn OR
               (local_PrevFlowLow AND local_PrevAlarmActive AND local_PrevAlarmAcked));

highHigh := NOT sensorOK;

local_PrevAckBtn := ackBtn;
local_PrevFlowLow := flowLow;
local_PrevAlarmActive := alarmActive;
local_PrevAlarmAcked := alarmAcked;

END_FUNCTION_BLOCK

(* ---- self-hard-02.candidate_01.st ---- *)
FUNCTION_BLOCK FB
VAR_INPUT
    startBtn : BOOL;
    abortBtn : BOOL;
    setpoint : REAL;
    pv : REAL;
    maxDuration : INT;
END_VAR
VAR_OUTPUT
    elapsed : INT;
    phase : INT;
    timeout : BOOL;
END_VAR
VAR
    localPrevStart : BOOL;
    localPrevPhase : INT;
    localPrevElapsed : INT;
    localPrevTimeout : BOOL;
    localRising : BOOL;
END_VAR

(* CONTRACT_RULES [] *)

(* ENGINEERING_CONTRACT
   - rising(startBtn): activated only when !abort; sets (phase, elapsed, timeout)=(1,0,FALSE).
   - abortBtn: highest same-scan priority; forces phase=9 and freezes elapsed/timeout.
   - running count: previous phase=1/2 increments elapsed by exactly 1 before phase/timeout evaluation.
   - timeout boundary: when elapsed >= maxDuration on this scan, set timeout=TRUE and phase=3.
   - heating boundary: not timed out, previous phase=1 and pv>=setpoint -> phase=2; phase=2 is retained.
   - frozen states: phase=0/3/9 retain phase, elapsed, and timeout until valid start or abort.
   - units: elapsed and maxDuration are integer scan counts; no TIME/LTIME or timer used.
   - start edge is consumed every scan, including same-scan abort, by updating localPrevStart.
*)

localRising := startBtn AND NOT localPrevStart;
localPrevPhase := phase;
localPrevElapsed := elapsed;
localPrevTimeout := timeout;

IF abortBtn THEN
    phase := 9;
    elapsed := localPrevElapsed;
    timeout := localPrevTimeout;
ELSIF localRising THEN
    phase := 1;
    elapsed := 0;
    timeout := FALSE;
ELSIF (localPrevPhase = 1) OR (localPrevPhase = 2) THEN
    elapsed := localPrevElapsed + 1;

    IF elapsed >= maxDuration THEN
        timeout := TRUE;
        phase := 3;
    ELSIF (localPrevPhase = 1) AND (pv >= setpoint) THEN
        timeout := FALSE;
        phase := 2;
    ELSIF localPrevPhase = 2 THEN
        timeout := FALSE;
        phase := 2;
    ELSE
        timeout := FALSE;
        phase := 1;
    END_IF;
ELSE
    phase := localPrevPhase;
    elapsed := localPrevElapsed;
    timeout := localPrevTimeout;
END_IF;

localPrevStart := startBtn;

END_FUNCTION_BLOCK

(* ---- self-hard-02.raw_candidate_01.st ---- *)
FUNCTION_BLOCK FB
VAR_INPUT
    startBtn : BOOL;
    abortBtn : BOOL;
    setpoint : REAL;
    pv : REAL;
    maxDuration : INT;
END_VAR
VAR_OUTPUT
    elapsed : INT;
    phase : INT;
    timeout : BOOL;
END_VAR
VAR
    localPrevStart : BOOL;
    localPrevPhase : INT;
    localPrevElapsed : INT;
    localPrevTimeout : BOOL;
    localRising : BOOL;
END_VAR

(* CONTRACT_RULES [] *)

(* ENGINEERING_CONTRACT
   - rising(startBtn): activated only when !abort; sets (phase, elapsed, timeout)=(1,0,FALSE).
   - abortBtn: highest same-scan priority; forces phase=9 and freezes elapsed/timeout.
   - running count: previous phase=1/2 increments elapsed by exactly 1 before phase/timeout evaluation.
   - timeout boundary: when elapsed >= maxDuration on this scan, set timeout=TRUE and phase=3.
   - heating boundary: not timed out, previous phase=1 and pv>=setpoint -> phase=2; phase=2 is retained.
   - frozen states: phase=0/3/9 retain phase, elapsed, and timeout until valid start or abort.
   - units: elapsed and maxDuration are integer scan counts; no TIME/LTIME or timer used.
   - start edge is consumed every scan, including same-scan abort, by updating localPrevStart.
*)

localRising := startBtn AND NOT localPrevStart;
localPrevPhase := phase;
localPrevElapsed := elapsed;
localPrevTimeout := timeout;

IF abortBtn THEN
    phase := 9;
    elapsed := localPrevElapsed;
    timeout := localPrevTimeout;
ELSIF localRising THEN
    phase := 1;
    elapsed := 0;
    timeout := FALSE;
ELSIF (localPrevPhase = 1) OR (localPrevPhase = 2) THEN
    elapsed := localPrevElapsed + 1;

    IF elapsed >= maxDuration THEN
        timeout := TRUE;
        phase := 3;
    ELSIF (localPrevPhase = 1) AND (pv >= setpoint) THEN
        timeout := FALSE;
        phase := 2;
    ELSIF localPrevPhase = 2 THEN
        timeout := FALSE;
        phase := 2;
    ELSE
        timeout := FALSE;
        phase := 1;
    END_IF
ELSE
    phase := localPrevPhase;
    elapsed := localPrevElapsed;
    timeout := localPrevTimeout;
END_IF

localPrevStart := startBtn;

END_FUNCTION_BLOCK

(* ---- self-hard-03.candidate_01.st ---- *)
(* CONTRACT_RULES [] *)
(* ENGINEERING_CONTRACT
  [PUB001] Capacity 8; inputs act only on FALSE->TRUE; initial count=0.
  [PUB002] popEn rising executes first: if count>0 shift fifo[1..7] left by one, decrement.
  [PUB003] pushEn rising executes second: if count<8 write fifo[count+1]=pushItem, increment.
  [PUB004] Same scan uses popped result; pop before push. Empty both => one item. Full both => replace one.
  [PUB005] count 0..8; full<=>count=8; empty<=>count=0.
  [PUB006] head=0 when empty, else head=fifo[1].
  [PUB007] fifo[1..count] remains compact in dequeue order; invalid tail unspecified.
  [PUB008] Retention: no successful operation preserves count and fifo[1..count]; push rejection preserves queue.
*)
FUNCTION_BLOCK FB
VAR_INPUT
    pushEn   : BOOL;
    pushItem : INT;
    popEn    : BOOL;
END_VAR
VAR_OUTPUT
    count : INT := 0;
    full  : BOOL := FALSE;
    empty : BOOL := TRUE;
    head  : INT := 0;
END_VAR
VAR_IN_OUT
    fifo : ARRAY[1..8] OF INT;
END_VAR
VAR
    local_push_prev : BOOL := FALSE;
    local_pop_prev  : BOOL := FALSE;
    local_push_rise : BOOL;
    local_pop_rise  : BOOL;
    local_count     : INT;
    local_i         : INT;
END_VAR

local_push_rise := pushEn AND NOT local_push_prev;
local_pop_rise  := popEn AND NOT local_pop_prev;

local_count := count;

IF local_pop_rise AND (local_count > 0) THEN
    FOR local_i := 1 TO 7 DO
        fifo[local_i] := fifo[local_i + 1];
    END_FOR;
    local_count := local_count - 1;
END_IF;

IF local_push_rise AND (local_count < 8) THEN
    fifo[local_count + 1] := pushItem;
    local_count := local_count + 1;
END_IF;

count := local_count;
full  := (count = 8);
empty := (count = 0);

IF count = 0 THEN
    head := 0;
ELSE
    head := fifo[1];
END_IF;

local_push_prev := pushEn;
local_pop_prev  := popEn;

END_FUNCTION_BLOCK

(* ---- self-hard-03.raw_candidate_01.st ---- *)
(* CONTRACT_RULES [] *)
(* ENGINEERING_CONTRACT
  [PUB001] Capacity 8; inputs act only on FALSE->TRUE; initial count=0.
  [PUB002] popEn rising executes first: if count>0 shift fifo[1..7] left by one, decrement.
  [PUB003] pushEn rising executes second: if count<8 write fifo[count+1]=pushItem, increment.
  [PUB004] Same scan uses popped result; pop before push. Empty both => one item. Full both => replace one.
  [PUB005] count 0..8; full<=>count=8; empty<=>count=0.
  [PUB006] head=0 when empty, else head=fifo[1].
  [PUB007] fifo[1..count] remains compact in dequeue order; invalid tail unspecified.
  [PUB008] Retention: no successful operation preserves count and fifo[1..count]; push rejection preserves queue.
*)
FUNCTION_BLOCK FB
VAR_INPUT
    pushEn   : BOOL;
    pushItem : INT;
    popEn    : BOOL;
END_VAR
VAR_OUTPUT
    count : INT := 0;
    full  : BOOL := FALSE;
    empty : BOOL := TRUE;
    head  : INT := 0;
END_VAR
VAR_IN_OUT
    fifo : ARRAY[1..8] OF INT;
END_VAR
VAR
    local_push_prev : BOOL := FALSE;
    local_pop_prev  : BOOL := FALSE;
    local_push_rise : BOOL;
    local_pop_rise  : BOOL;
    local_count     : INT;
    local_i         : INT;
END_VAR

local_push_rise := pushEn AND NOT local_push_prev;
local_pop_rise  := popEn AND NOT local_pop_prev;

local_count := count;

IF local_pop_rise AND (local_count > 0) THEN
    FOR local_i := 1 TO 7 DO
        fifo[local_i] := fifo[local_i + 1];
    END_FOR;
    local_count := local_count - 1;
END_IF;

IF local_push_rise AND (local_count < 8) THEN
    fifo[local_count + 1] := pushItem;
    local_count := local_count + 1;
END_IF;

count := local_count;
full  := (count = 8);
empty := (count = 0);

IF count = 0 THEN
    head := 0;
ELSE
    head := fifo[1];
END_IF;

local_push_prev := pushEn;
local_pop_prev  := popEn;

END_FUNCTION_BLOCK

(* ---- self-hard-04.candidate_01.st ---- *)
FUNCTION_BLOCK FB
VAR_INPUT
    demand : INT;
    runHours : ARRAY[1..5] OF LINT;
    rotated : BOOL;
END_VAR
VAR_OUTPUT
    leadPump : INT;
    lagPump : INT;
    runningCount : INT;
END_VAR
VAR
    local_clamped : INT := 0;
    local_minPump : INT := 0;
    local_candidateLag : INT := 0;
    local_prevLead : INT := 0;
    local_prevLag : INT := 0;
    local_prevRunningCount : INT := 0;
    local_leadChanged : BOOL := FALSE;
    local_countRise : BOOL := FALSE;
    tmp_i : INT := 0;
END_VAR

(* ENGINEERING_CONTRACT
   runningCount: clamps demand to 0..5 each scan; demand<=0 also clears selections (PUB001/S1/S5).
   leadPump activation: positive restart/init selects global min by (hours,pump#).
   leadPump hold: level rotated swaps only when previous valid lead-min>50h; otherwise holds; no rotated holds (PUB002/S3/S6/S7).
   lead/lag reset: demand=0 sets both 0 same scan (S4).
   lagPump activation/reselect: only initial, clamped demand rise, or lead change; choose min excluding new lead (PUB003/S8).
   lagPump hold: while demand>=2, lead unchanged and count not rising, lag remains previous (S9).
   Same-scan order: clamp->lead->lag; all hours LINT, threshold strict >50; array slots 1..5 only.
*)

(* CONTRACT_RULES [] *)

IF demand < 0 THEN
    local_clamped := 0;
ELSIF demand > 5 THEN
    local_clamped := 5;
ELSE
    local_clamped := demand;
END_IF;

runningCount := local_clamped;

IF local_clamped = 0 THEN
    leadPump := 0;
    lagPump := 0;
ELSE
    local_minPump := 1;
    FOR tmp_i := 2 TO 5 DO
        IF runHours[tmp_i] < runHours[local_minPump] THEN
            local_minPump := tmp_i;
        END_IF;
    END_FOR;

    IF (local_prevLead < 1) OR (local_prevLead > 5) THEN
        leadPump := local_minPump;
    ELSIF NOT rotated THEN
        leadPump := local_prevLead;
    ELSIF (runHours[local_prevLead] - runHours[local_minPump]) > 50 THEN
        leadPump := local_minPump;
    ELSE
        leadPump := local_prevLead;
    END_IF;

    IF local_clamped < 2 THEN
        lagPump := 0;
    ELSE
        local_leadChanged := (leadPump <> local_prevLead);
        local_countRise := local_clamped > local_prevRunningCount;

        IF local_leadChanged OR local_countRise THEN
            local_candidateLag := 0;
            FOR tmp_i := 1 TO 5 DO
                IF tmp_i <> leadPump THEN
                    IF local_candidateLag = 0 THEN
                        local_candidateLag := tmp_i;
                    ELSIF runHours[tmp_i] < runHours[local_candidateLag] THEN
                        local_candidateLag := tmp_i;
                    END_IF;
                END_IF;
            END_FOR;
            lagPump := local_candidateLag;
        ELSE
            lagPump := local_prevLag;
        END_IF;
    END_IF;
END_IF;

local_prevLead := leadPump;
local_prevLag := lagPump;
local_prevRunningCount := local_clamped;

END_FUNCTION_BLOCK

(* ---- self-hard-04.raw_candidate_01.st ---- *)
FUNCTION_BLOCK FB
VAR_INPUT
    demand : INT;
    runHours : ARRAY[1..5] OF LINT;
    rotated : BOOL;
END_VAR
VAR_OUTPUT
    leadPump : INT;
    lagPump : INT;
    runningCount : INT;
END_VAR
VAR
    local_clamped : INT := 0;
    local_minPump : INT := 0;
    local_candidateLag : INT := 0;
    local_prevLead : INT := 0;
    local_prevLag : INT := 0;
    local_prevRunningCount : INT := 0;
    local_leadChanged : BOOL := FALSE;
    local_countRise : BOOL := FALSE;
    tmp_i : INT := 0;
END_VAR

(* ENGINEERING_CONTRACT
   runningCount: clamps demand to 0..5 each scan; demand<=0 also clears selections (PUB001/S1/S5).
   leadPump activation: positive restart/init selects global min by (hours,pump#).
   leadPump hold: level rotated swaps only when previous valid lead-min>50h; otherwise holds; no rotated holds (PUB002/S3/S6/S7).
   lead/lag reset: demand=0 sets both 0 same scan (S4).
   lagPump activation/reselect: only initial, clamped demand rise, or lead change; choose min excluding new lead (PUB003/S8).
   lagPump hold: while demand>=2, lead unchanged and count not rising, lag remains previous (S9).
   Same-scan order: clamp->lead->lag; all hours LINT, threshold strict >50; array slots 1..5 only.
*)

(* CONTRACT_RULES [] *)

IF demand < 0 THEN
    local_clamped := 0;
ELSIF demand > 5 THEN
    local_clamped := 5;
ELSE
    local_clamped := demand;
END_IF;

runningCount := local_clamped;

IF local_clamped = 0 THEN
    leadPump := 0;
    lagPump := 0;
ELSE
    local_minPump := 1;
    FOR tmp_i := 2 TO 5 DO
        IF runHours[tmp_i] < runHours[local_minPump] THEN
            local_minPump := tmp_i;
        END_IF;
    END_FOR;

    IF (local_prevLead < 1) OR (local_prevLead > 5) THEN
        leadPump := local_minPump;
    ELSIF NOT rotated THEN
        leadPump := local_prevLead;
    ELSIF (runHours[local_prevLead] - runHours[local_minPump]) > 50 THEN
        leadPump := local_minPump;
    ELSE
        leadPump := local_prevLead;
    END_IF;

    IF local_clamped < 2 THEN
        lagPump := 0;
    ELSE
        local_leadChanged := (leadPump <> local_prevLead);
        local_countRise := local_clamped > local_prevRunningCount;

        IF local_leadChanged OR local_countRise THEN
            local_candidateLag := 0;
            FOR tmp_i := 1 TO 5 DO
                IF tmp_i <> leadPump THEN
                    IF local_candidateLag = 0 THEN
                        local_candidateLag := tmp_i;
                    ELSIF runHours[tmp_i] < runHours[local_candidateLag] THEN
                        local_candidateLag := tmp_i;
                    END_IF;
                END_IF;
            END_FOR;
            lagPump := local_candidateLag;
        ELSE
            lagPump := local_prevLag;
        END_IF;
    END_IF;
END_IF;

local_prevLead := leadPump;
local_prevLag := lagPump;
local_prevRunningCount := local_clamped;

END_FUNCTION_BLOCK

(* ---- self-hard-05.candidate_01.st ---- *)
FUNCTION_BLOCK FB
VAR_INPUT
    runRequest : BOOL;
    flameOK : BOOL;
    o2Valid : BOOL;
    o2PV : REAL;
    baseAir : REAL;
    resetBtn : BOOL;
END_VAR
VAR_OUTPUT
    fuelPermit : BOOL;
    trimEnable : BOOL;
    airTrim : REAL;
    airCommand : REAL;
    tripLatched : BOOL;
    o2Fault : BOOL;
END_VAR
VAR
    local_resetEdge : R_TRIG;
    tmp_resetRising : BOOL;
    tmp_rawTrim : REAL;
    tmp_rawAir : REAL;
END_VAR

(* ENGINEERING_CONTRACT
tripLatched: set same scan when runRequest & !flameOK; holds; reset only resetBtn rising with !runRequest & !flameOK (PUB001/PUB002).
fuelPermit: runRequest & flameOK & !tripLatched, evaluated after trip update (PUB003).
o2Fault: !o2Valid OR o2PV<0.0 OR o2PV>21.0; combinational, does not cut fuel (PUB005).
trimEnable: fuelPermit & !o2Fault; combinational after fuel/fault update (PUB004/PUB008).
airTrim: if trimEnable then clamp(2.0*(2.0-o2PV),-10.0,10.0), else 0.0; units % (PUB004/PUB006).
airCommand: if fuelPermit then clamp(baseAir+airTrim,0.0,100.0), else 0.0; baseAir itself not bounded (PUB006).
R_TRIG evaluated before state equations; held resetBtn has no repeated effect; units: o2PV/baseAir/airTrim/airCommand %.
*)
(* CONTRACT_RULES [] *)

local_resetEdge(CLK := resetBtn);
tmp_resetRising := local_resetEdge.Q;

tripLatched := (runRequest AND NOT flameOK)
    OR (tripLatched AND NOT (tmp_resetRising AND NOT runRequest AND NOT flameOK));

fuelPermit := runRequest AND flameOK AND NOT tripLatched;

o2Fault := (NOT o2Valid) OR (o2PV < 0.0) OR (o2PV > 21.0);

trimEnable := fuelPermit AND NOT o2Fault;

IF trimEnable THEN
    tmp_rawTrim := 2.0 * (2.0 - o2PV);
    IF tmp_rawTrim > 10.0 THEN
        airTrim := 10.0;
    ELSIF tmp_rawTrim < -10.0 THEN
        airTrim := -10.0;
    ELSE
        airTrim := tmp_rawTrim;
    END_IF;
ELSE
    airTrim := 0.0;
END_IF;

IF fuelPermit THEN
    tmp_rawAir := baseAir + airTrim;
    IF tmp_rawAir > 100.0 THEN
        airCommand := 100.0;
    ELSIF tmp_rawAir < 0.0 THEN
        airCommand := 0.0;
    ELSE
        airCommand := tmp_rawAir;
    END_IF;
ELSE
    airCommand := 0.0;
END_IF;

END_FUNCTION_BLOCK

(* ---- self-hard-05.raw_candidate_01.st ---- *)
FUNCTION_BLOCK FB
VAR_INPUT
    runRequest : BOOL;
    flameOK : BOOL;
    o2Valid : BOOL;
    o2PV : REAL;
    baseAir : REAL;
    resetBtn : BOOL;
END_VAR
VAR_OUTPUT
    fuelPermit : BOOL;
    trimEnable : BOOL;
    airTrim : REAL;
    airCommand : REAL;
    tripLatched : BOOL;
    o2Fault : BOOL;
END_VAR
VAR
    local_resetEdge : R_TRIG;
    tmp_resetRising : BOOL;
    tmp_rawTrim : REAL;
    tmp_rawAir : REAL;
END_VAR

(* ENGINEERING_CONTRACT
tripLatched: set same scan when runRequest & !flameOK; holds; reset only resetBtn rising with !runRequest & !flameOK (PUB001/PUB002).
fuelPermit: runRequest & flameOK & !tripLatched, evaluated after trip update (PUB003).
o2Fault: !o2Valid OR o2PV<0.0 OR o2PV>21.0; combinational, does not cut fuel (PUB005).
trimEnable: fuelPermit & !o2Fault; combinational after fuel/fault update (PUB004/PUB008).
airTrim: if trimEnable then clamp(2.0*(2.0-o2PV),-10.0,10.0), else 0.0; units % (PUB004/PUB006).
airCommand: if fuelPermit then clamp(baseAir+airTrim,0.0,100.0), else 0.0; baseAir itself not bounded (PUB006).
R_TRIG evaluated before state equations; held resetBtn has no repeated effect; units: o2PV/baseAir/airTrim/airCommand %.
*)
(* CONTRACT_RULES [] *)

local_resetEdge(CLK := resetBtn);
tmp_resetRising := local_resetEdge.Q;

tripLatched := (runRequest AND NOT flameOK)
    OR (tripLatched AND NOT (tmp_resetRising AND NOT runRequest AND NOT flameOK));

fuelPermit := runRequest AND flameOK AND NOT tripLatched;

o2Fault := (NOT o2Valid) OR (o2PV < 0.0) OR (o2PV > 21.0);

trimEnable := fuelPermit AND NOT o2Fault;

IF trimEnable THEN
    tmp_rawTrim := 2.0 * (2.0 - o2PV);
    IF tmp_rawTrim > 10.0 THEN
        airTrim := 10.0;
    ELSIF tmp_rawTrim < -10.0 THEN
        airTrim := -10.0;
    ELSE
        airTrim := tmp_rawTrim;
    END_IF;
ELSE
    airTrim := 0.0;
END_IF;

IF fuelPermit THEN
    tmp_rawAir := baseAir + airTrim;
    IF tmp_rawAir > 100.0 THEN
        airCommand := 100.0;
    ELSIF tmp_rawAir < 0.0 THEN
        airCommand := 0.0;
    ELSE
        airCommand := tmp_rawAir;
    END_IF;
ELSE
    airCommand := 0.0;
END_IF;

END_FUNCTION_BLOCK

(* ---- self-hard-06.candidate_01.st ---- *)
FUNCTION_BLOCK FB
VAR_INPUT
    runRequest : BOOL;
    pressure : REAL;
    pressureValid : BOOL;
    fuelFlow : REAL;
    steamFlow : REAL;
    outletCmd : INT;
    outletFeedback : INT;
    resetBtn : BOOL;
END_VAR
VAR_OUTPUT
    tripLatched : BOOL;
    fuelPermit : BOOL;
    currentCauseMask : WORD;
    latchedCauseMask : WORD;
    diagnosticActive : BOOL;
END_VAR
VAR
    tmp_resetPrev : BOOL;
    tmp_resetRising : BOOL;
    tmp_legalReset : BOOL;
    tmp_overpressure : BOOL;
    tmp_valvePred : BOOL;
    tmp_valveStuck : BOOL;
    tmp_combustion : BOOL;
    tmp_tripCondition : BOOL;
    tmp_tripNew : BOOL;
    tmp_previousLatched : WORD;
    tmp_stuckCycles : UINT;
END_VAR

(* ENGINEERING_CONTRACT
  tripLatched: set same scan by run & (!pressureValid OR pressure >= 4500.0); retained; cleared only legal reset edge (!run & valid & p <= 4200.0). PUB004-PUB007/PUB012.
  fuelPermit: run & NOT tripLatched. diagnosticActive: currentCauseMask <> 0. PUB021-PUB023.
  currentCauseMask low nibble: !run = 0; invalid = 1; valid overpressure = 2/4/6/8; valid below 4500 = 0. PUB024-PUB035.
  valve bit: 3 consecutive true scans of valid-overpressure valve criterion; any false criterion scan clears the cycle counter. PUB034.
  latchedCauseMask: when final tripLatched is true, old footprint OR current mask; zero when not tripped or on legal reset. PUB036.
  REAL boundaries inclusive: trip >= 4500.0, reset <= 4200.0, fuel >= 4.0, steam <= 10.0; cycles not seconds. PUB027/PUB040.
*)

(* CONTRACT_RULES [] *)

tmp_resetRising := resetBtn AND NOT tmp_resetPrev;
tmp_legalReset := tmp_resetRising AND NOT runRequest AND pressureValid AND (pressure <= 4200.0);

tmp_overpressure := runRequest AND pressureValid AND (pressure >= 4500.0);
tmp_valvePred := runRequest AND pressureValid AND (pressure >= 4500.0)
                 AND (outletCmd >= 50) AND (outletFeedback <= 10);
tmp_combustion := (fuelFlow >= 4.0) AND (steamFlow <= 10.0);

IF tmp_valvePred THEN
    IF tmp_stuckCycles < UINT#3 THEN
        tmp_stuckCycles := tmp_stuckCycles + UINT#1;
    END_IF;
ELSE
    tmp_stuckCycles := UINT#0;
END_IF;

tmp_valveStuck := tmp_stuckCycles >= UINT#3;

IF NOT runRequest THEN
    currentCauseMask := WORD#0;
ELSIF NOT pressureValid THEN
    currentCauseMask := WORD#1;
ELSIF pressure >= 4500.0 THEN
    IF tmp_valveStuck AND tmp_combustion THEN
        currentCauseMask := WORD#6;
    ELSIF tmp_valveStuck THEN
        currentCauseMask := WORD#2;
    ELSIF tmp_combustion THEN
        currentCauseMask := WORD#4;
    ELSE
        currentCauseMask := WORD#8;
    END_IF;
ELSE
    currentCauseMask := WORD#0;
END_IF;

tmp_tripCondition := runRequest AND (NOT pressureValid OR (pressure >= 4500.0));
tmp_previousLatched := latchedCauseMask;

tmp_tripNew := tripLatched;
IF tmp_legalReset THEN
    tmp_tripNew := FALSE;
ELSIF tmp_tripCondition THEN
    tmp_tripNew := TRUE;
END_IF;

IF tmp_legalReset THEN
    latchedCauseMask := WORD#0;
ELSIF tmp_tripNew THEN
    latchedCauseMask := tmp_previousLatched OR currentCauseMask;
ELSE
    latchedCauseMask := WORD#0;
END_IF;

tripLatched := tmp_tripNew;
fuelPermit := runRequest AND NOT tripLatched;
diagnosticActive := currentCauseMask <> WORD#0;

tmp_resetPrev := resetBtn;
END_FUNCTION_BLOCK

(* ---- self-hard-06.raw_candidate_01.st ---- *)
FUNCTION_BLOCK FB
VAR_INPUT
    runRequest : BOOL;
    pressure : REAL;
    pressureValid : BOOL;
    fuelFlow : REAL;
    steamFlow : REAL;
    outletCmd : INT;
    outletFeedback : INT;
    resetBtn : BOOL;
END_VAR
VAR_OUTPUT
    tripLatched : BOOL;
    fuelPermit : BOOL;
    currentCauseMask : WORD;
    latchedCauseMask : WORD;
    diagnosticActive : BOOL;
END_VAR
VAR
    tmp_resetPrev : BOOL;
    tmp_resetRising : BOOL;
    tmp_legalReset : BOOL;
    tmp_overpressure : BOOL;
    tmp_valvePred : BOOL;
    tmp_valveStuck : BOOL;
    tmp_combustion : BOOL;
    tmp_tripCondition : BOOL;
    tmp_tripNew : BOOL;
    tmp_previousLatched : WORD;
    tmp_stuckCycles : UINT;
END_VAR

(* ENGINEERING_CONTRACT
  tripLatched: set same scan by run & (!pressureValid OR pressure >= 4500.0); retained; cleared only legal reset edge (!run & valid & p <= 4200.0). PUB004-PUB007/PUB012.
  fuelPermit: run & NOT tripLatched. diagnosticActive: currentCauseMask <> 0. PUB021-PUB023.
  currentCauseMask low nibble: !run = 0; invalid = 1; valid overpressure = 2/4/6/8; valid below 4500 = 0. PUB024-PUB035.
  valve bit: 3 consecutive true scans of valid-overpressure valve criterion; any false criterion scan clears the cycle counter. PUB034.
  latchedCauseMask: when final tripLatched is true, old footprint OR current mask; zero when not tripped or on legal reset. PUB036.
  REAL boundaries inclusive: trip >= 4500.0, reset <= 4200.0, fuel >= 4.0, steam <= 10.0; cycles not seconds. PUB027/PUB040.
*)

(* CONTRACT_RULES [] *)

tmp_resetRising := resetBtn AND NOT tmp_resetPrev;
tmp_legalReset := tmp_resetRising AND NOT runRequest AND pressureValid AND (pressure <= 4200.0);

tmp_overpressure := runRequest AND pressureValid AND (pressure >= 4500.0);
tmp_valvePred := runRequest AND pressureValid AND (pressure >= 4500.0)
                 AND (outletCmd >= 50) AND (outletFeedback <= 10);
tmp_combustion := (fuelFlow >= 4.0) AND (steamFlow <= 10.0);

IF tmp_valvePred THEN
    IF tmp_stuckCycles < UINT#3 THEN
        tmp_stuckCycles := tmp_stuckCycles + UINT#1;
    END_IF;
ELSE
    tmp_stuckCycles := UINT#0;
END_IF;

tmp_valveStuck := tmp_stuckCycles >= UINT#3;

IF NOT runRequest THEN
    currentCauseMask := WORD#0;
ELSIF NOT pressureValid THEN
    currentCauseMask := WORD#1;
ELSIF pressure >= 4500.0 THEN
    IF tmp_valveStuck AND tmp_combustion THEN
        currentCauseMask := WORD#6;
    ELSIF tmp_valveStuck THEN
        currentCauseMask := WORD#2;
    ELSIF tmp_combustion THEN
        currentCauseMask := WORD#4;
    ELSE
        currentCauseMask := WORD#8;
    END_IF;
ELSE
    currentCauseMask := WORD#0;
END_IF;

tmp_tripCondition := runRequest AND (NOT pressureValid OR (pressure >= 4500.0));
tmp_previousLatched := latchedCauseMask;

tmp_tripNew := tripLatched;
IF tmp_legalReset THEN
    tmp_tripNew := FALSE;
ELSIF tmp_tripCondition THEN
    tmp_tripNew := TRUE;
END_IF;

IF tmp_legalReset THEN
    latchedCauseMask := WORD#0;
ELSIF tmp_tripNew THEN
    latchedCauseMask := tmp_previousLatched OR currentCauseMask;
ELSE
    latchedCauseMask := WORD#0;
END_IF;

tripLatched := tmp_tripNew;
fuelPermit := runRequest AND NOT tripLatched;
diagnosticActive := currentCauseMask <> WORD#0;

tmp_resetPrev := resetBtn;
END_FUNCTION_BLOCK

(* ---- self-hard-07.candidate_01.st ---- *)
FUNCTION_BLOCK FB
VAR_INPUT
    mode : INT;
    resetBtn : BOOL;
    scanSeconds : REAL;
    tempSP : REAL;
    tempPV : REAL;
    flowPV : REAL;
    manualFlowSP : REAL;
    manualValve : REAL;
END_VAR
VAR_OUTPUT
    flowSP : REAL;
    valveCommand : REAL;
    fault : BOOL;
    normalMode : BOOL;
END_VAR
VAR
    accT : REAL;
    accF : REAL;
    eT : REAL;
    eF : REAL;
    raw : REAL;
    local_hasPrev : BOOL;
    local_prevMode : INT;
    local_prevReset : BOOL;
    local_modeChanged : BOOL;
    local_resetEdge : BOOL;
END_VAR

(* ENGINEERING_CONTRACT
   flowSP: bounded 0..50 t/h (S1). valveCommand: bounded 0..100 % (S2).
   fault: invalid mode/scanSeconds -> manual outputs, no PI, normalMode false (PUB006,S3,S10).
   reset edge: manual outputs, no PI, edge memory; hold does not repeat (PUB005,S4).
   transition: to mode 1/0 flowSP=manual and valve holds; to mode 2 both hold; normal false (PUB004,S7,S8).
   normalMode: prior scan exists, mode stable, no fault, no reset edge (S11).
   normal PI: cascade outer then inner; accT/accF back-calculated from clamped outputs (PUB003,S13,S14).
   manual normal: both outputs follow manual values (S5); auto flowSP=manual (S6).
   same-scan priority: reset > fault > first scan > mode change > normal; fault still reported on reset scan.
*)

(* CONTRACT_RULES [] *)

eT := tempSP - tempPV;

fault := (mode < 0) OR (mode > 2) OR (scanSeconds <= 0.0) OR (scanSeconds > 10.0);

local_resetEdge := resetBtn AND NOT local_prevReset;
local_modeChanged := local_hasPrev AND (mode <> local_prevMode);

IF local_resetEdge THEN
    flowSP := manualFlowSP;
    valveCommand := manualValve;
ELSIF fault THEN
    flowSP := manualFlowSP;
    valveCommand := manualValve;
ELSIF NOT local_hasPrev THEN
    flowSP := manualFlowSP;
    valveCommand := manualValve;
ELSIF local_modeChanged THEN
    IF mode = 2 THEN
        flowSP := flowSP;
    ELSE
        flowSP := manualFlowSP;
    END_IF;
    valveCommand := valveCommand;
ELSE
    IF mode = 0 THEN
        flowSP := manualFlowSP;
        valveCommand := manualValve;
    ELSIF mode = 1 THEN
        flowSP := manualFlowSP;
        eF := flowSP - flowPV;
        raw := accF + 2.0 * eF + 0.5 * eF * scanSeconds;
        valveCommand := LIMIT(0.0, raw, 100.0);
    ELSIF mode = 2 THEN
        raw := accT + 1.0 * eT + 0.2 * eT * scanSeconds;
        flowSP := LIMIT(0.0, raw, 50.0);

        eF := flowSP - flowPV;
        raw := accF + 2.0 * eF + 0.5 * eF * scanSeconds;
        valveCommand := LIMIT(0.0, raw, 100.0);
    END_IF;
END_IF;

eF := flowSP - flowPV;
accT := flowSP - 1.0 * eT;
accF := valveCommand - 2.0 * eF;

normalMode := local_hasPrev AND (mode = local_prevMode) AND NOT fault AND NOT local_resetEdge;

local_prevMode := mode;
local_prevReset := resetBtn;
local_hasPrev := TRUE;

END_FUNCTION_BLOCK

(* ---- self-hard-07.raw_candidate_01.st ---- *)
FUNCTION_BLOCK FB
VAR_INPUT
    mode : INT;
    resetBtn : BOOL;
    scanSeconds : REAL;
    tempSP : REAL;
    tempPV : REAL;
    flowPV : REAL;
    manualFlowSP : REAL;
    manualValve : REAL;
END_VAR
VAR_OUTPUT
    flowSP : REAL;
    valveCommand : REAL;
    fault : BOOL;
    normalMode : BOOL;
END_VAR
VAR
    accT : REAL;
    accF : REAL;
    eT : REAL;
    eF : REAL;
    raw : REAL;
    local_hasPrev : BOOL;
    local_prevMode : INT;
    local_prevReset : BOOL;
    local_modeChanged : BOOL;
    local_resetEdge : BOOL;
END_VAR

(* ENGINEERING_CONTRACT
   flowSP: bounded 0..50 t/h (S1). valveCommand: bounded 0..100 % (S2).
   fault: invalid mode/scanSeconds -> manual outputs, no PI, normalMode false (PUB006,S3,S10).
   reset edge: manual outputs, no PI, edge memory; hold does not repeat (PUB005,S4).
   transition: to mode 1/0 flowSP=manual and valve holds; to mode 2 both hold; normal false (PUB004,S7,S8).
   normalMode: prior scan exists, mode stable, no fault, no reset edge (S11).
   normal PI: cascade outer then inner; accT/accF back-calculated from clamped outputs (PUB003,S13,S14).
   manual normal: both outputs follow manual values (S5); auto flowSP=manual (S6).
   same-scan priority: reset > fault > first scan > mode change > normal; fault still reported on reset scan.
*)

(* CONTRACT_RULES [] *)

eT := tempSP - tempPV;

fault := (mode < 0) OR (mode > 2) OR (scanSeconds <= 0.0) OR (scanSeconds > 10.0);

local_resetEdge := resetBtn AND NOT local_prevReset;
local_modeChanged := local_hasPrev AND (mode <> local_prevMode);

IF local_resetEdge THEN
    flowSP := manualFlowSP;
    valveCommand := manualValve;
ELSIF fault THEN
    flowSP := manualFlowSP;
    valveCommand := manualValve;
ELSIF NOT local_hasPrev THEN
    flowSP := manualFlowSP;
    valveCommand := manualValve;
ELSIF local_modeChanged THEN
    IF mode = 2 THEN
        flowSP := flowSP;
    ELSE
        flowSP := manualFlowSP;
    END_IF;
    valveCommand := valveCommand;
ELSE
    IF mode = 0 THEN
        flowSP := manualFlowSP;
        valveCommand := manualValve;
    ELSIF mode = 1 THEN
        flowSP := manualFlowSP;
        eF := flowSP - flowPV;
        raw := accF + 2.0 * eF + 0.5 * eF * scanSeconds;
        valveCommand := LIMIT(0.0, raw, 100.0);
    ELSIF mode = 2 THEN
        raw := accT + 1.0 * eT + 0.2 * eT * scanSeconds;
        flowSP := LIMIT(0.0, raw, 50.0);

        eF := flowSP - flowPV;
        raw := accF + 2.0 * eF + 0.5 * eF * scanSeconds;
        valveCommand := LIMIT(0.0, raw, 100.0);
    END_IF;
END_IF;

eF := flowSP - flowPV;
accT := flowSP - 1.0 * eT;
accF := valveCommand - 2.0 * eF;

normalMode := local_hasPrev AND (mode = local_prevMode) AND NOT fault AND NOT local_resetEdge;

local_prevMode := mode;
local_prevReset := resetBtn;
local_hasPrev := TRUE;

END_FUNCTION_BLOCK

(* ---- self-medium-01.candidate_01.st ---- *)
TYPE ST_Recipe :
STRUCT
    recipeID : INT;
    totalRatio : REAL;
    temperature : REAL;
END_STRUCT
END_TYPE;

FUNCTION_BLOCK FB
VAR_INPUT
    recipe : ARRAY[1..8] OF ST_Recipe;
    selSlot : INT;
    loadCmd : BOOL;
    running : BOOL;
END_VAR
VAR_OUTPUT
    valid : BOOL;
    loadedID : INT;
END_VAR
VAR
    tmp_cmd_was_high : BOOL := FALSE;
    tmp_rising : BOOL;
    tmp_prev_valid : BOOL;
    tmp_prev_loaded : INT;
END_VAR

(* ENGINEERING_CONTRACT
- valid activates only on !running AND rising(loadCmd); otherwise it holds the prior value.
- valid TRUE iff selSlot is 1..8 and the selected slot is non-empty with totalRatio in [99.0,101.0] and temperature in [30.0,180.0]; otherwise FALSE.
- loadedID is set to the selected recipeID on a valid load and to 0 on an invalid load; otherwise it holds the prior value.
- running TRUE suppresses loading and preserves prior valid and loadedID (N10-S4,S9).
- recipe[selSlot] is dereferenced only after bounds validation; a held loadCmd does not retrigger (S5,S6).
*)

(* CONTRACT_RULES [] *)

tmp_rising := loadCmd AND NOT tmp_cmd_was_high;
tmp_prev_valid := valid;
tmp_prev_loaded := loadedID;

IF (NOT running) AND tmp_rising THEN
    IF (selSlot >= 1) AND (selSlot <= 8) THEN
        IF (recipe[selSlot].recipeID <> 0)
           AND (recipe[selSlot].totalRatio >= 99.0)
           AND (recipe[selSlot].totalRatio <= 101.0)
           AND (recipe[selSlot].temperature >= 30.0)
           AND (recipe[selSlot].temperature <= 180.0) THEN
            valid := TRUE;
            loadedID := recipe[selSlot].recipeID;
        ELSE
            valid := FALSE;
            loadedID := 0;
        END_IF;
    ELSE
        valid := FALSE;
        loadedID := 0;
    END_IF;
ELSE
    valid := tmp_prev_valid;
    loadedID := tmp_prev_loaded;
END_IF;

tmp_cmd_was_high := loadCmd;
END_FUNCTION_BLOCK

(* ---- self-medium-01.raw_candidate_01.st ---- *)
TYPE ST_Recipe :
STRUCT
    recipeID : INT;
    totalRatio : REAL;
    temperature : REAL;
END_STRUCT
END_TYPE

FUNCTION_BLOCK FB
VAR_INPUT
    recipe : ARRAY[1..8] OF ST_Recipe;
    selSlot : INT;
    loadCmd : BOOL;
    running : BOOL;
END_VAR
VAR_OUTPUT
    valid : BOOL;
    loadedID : INT;
END_VAR
VAR
    tmp_cmd_was_high : BOOL := FALSE;
    tmp_rising : BOOL;
    tmp_prev_valid : BOOL;
    tmp_prev_loaded : INT;
END_VAR

(* ENGINEERING_CONTRACT
- valid activates only on !running AND rising(loadCmd); otherwise it holds the prior value.
- valid TRUE iff selSlot is 1..8 and the selected slot is non-empty with totalRatio in [99.0,101.0] and temperature in [30.0,180.0]; otherwise FALSE.
- loadedID is set to the selected recipeID on a valid load and to 0 on an invalid load; otherwise it holds the prior value.
- running TRUE suppresses loading and preserves prior valid and loadedID (N10-S4,S9).
- recipe[selSlot] is dereferenced only after bounds validation; a held loadCmd does not retrigger (S5,S6).
*)

(* CONTRACT_RULES [] *)

tmp_rising := loadCmd AND NOT tmp_cmd_was_high;
tmp_prev_valid := valid;
tmp_prev_loaded := loadedID;

IF (NOT running) AND tmp_rising THEN
    IF (selSlot >= 1) AND (selSlot <= 8) THEN
        IF (recipe[selSlot].recipeID <> 0)
           AND (recipe[selSlot].totalRatio >= 99.0)
           AND (recipe[selSlot].totalRatio <= 101.0)
           AND (recipe[selSlot].temperature >= 30.0)
           AND (recipe[selSlot].temperature <= 180.0) THEN
            valid := TRUE;
            loadedID := recipe[selSlot].recipeID;
        ELSE
            valid := FALSE;
            loadedID := 0;
        END_IF;
    ELSE
        valid := FALSE;
        loadedID := 0;
    END_IF;
ELSE
    valid := tmp_prev_valid;
    loadedID := tmp_prev_loaded;
END_IF;

tmp_cmd_was_high := loadCmd;
END_FUNCTION_BLOCK

(* ---- self-medium-02.candidate_01.st ---- *)
FUNCTION_BLOCK FB
VAR_INPUT
    enable : BOOL;
    rawValue : REAL;
END_VAR
VAR_OUTPUT
    filteredValue : REAL;
    windowFull : BOOL;
    sampleCount : INT;
END_VAR
VAR
    tmp_buffer : ARRAY[0..7] OF REAL;
    tmp_count : INT := 0;
    tmp_write_index : INT := 0;
    tmp_sum : REAL := 0.0;
    tmp_i : INT := 0;
END_VAR

(* ENGINEERING_CONTRACT
- filteredValue: recomputed every enabled scan after push; disabled scan retains last mean (PUB005, PUB010).
- sampleCount: 0..8, increments while enabled and <8, holds at 8, resets same scan when disabled (PUB008, PUB010).
- windowFull: TRUE exactly when tmp_count=8; held until disable resets FALSE (PUB009, PUB010).
- FIFO: non-full uses actual count, no zero padding; full replaces oldest (PUB006, PUB007).
- new period: independent count; first enabled sample outputs raw, second outputs two-sample mean (PUB011, S6-S7).
- unspecified: disable ignores rawValue; stored array bits may remain but count defines validity.
*)

IF enable THEN
    IF tmp_count < 8 THEN
        tmp_buffer[tmp_count] := rawValue;
        tmp_count := tmp_count + 1;
        IF tmp_count < 8 THEN
            tmp_write_index := tmp_count;
        ELSE
            tmp_write_index := 0;
        END_IF;
    ELSE
        tmp_buffer[tmp_write_index] := rawValue;
        tmp_write_index := tmp_write_index + 1;
        IF tmp_write_index > 7 THEN
            tmp_write_index := 0;
        END_IF;
    END_IF;

    tmp_sum := 0.0;
    FOR tmp_i := 0 TO tmp_count - 1 DO
        tmp_sum := tmp_sum + tmp_buffer[tmp_i];
    END_FOR;

    IF tmp_count > 0 THEN
        filteredValue := tmp_sum / INT_TO_REAL(tmp_count);
    END_IF;

    sampleCount := tmp_count;
    windowFull := (tmp_count = 8);
ELSE
    tmp_count := 0;
    tmp_write_index := 0;
    sampleCount := 0;
    windowFull := FALSE;
END_IF;

(* CONTRACT_RULES [] *)

END_FUNCTION_BLOCK

(* ---- self-medium-02.raw_candidate_01.st ---- *)
FUNCTION_BLOCK FB
VAR_INPUT
    enable : BOOL;
    rawValue : REAL;
END_VAR
VAR_OUTPUT
    filteredValue : REAL;
    windowFull : BOOL;
    sampleCount : INT;
END_VAR
VAR
    tmp_buffer : ARRAY[0..7] OF REAL;
    tmp_count : INT := 0;
    tmp_write_index : INT := 0;
    tmp_sum : REAL := 0.0;
    tmp_i : INT := 0;
END_VAR

(* ENGINEERING_CONTRACT
- filteredValue: recomputed every enabled scan after push; disabled scan retains last mean (PUB005, PUB010).
- sampleCount: 0..8, increments while enabled and <8, holds at 8, resets same scan when disabled (PUB008, PUB010).
- windowFull: TRUE exactly when tmp_count=8; held until disable resets FALSE (PUB009, PUB010).
- FIFO: non-full uses actual count, no zero padding; full replaces oldest (PUB006, PUB007).
- new period: independent count; first enabled sample outputs raw, second outputs two-sample mean (PUB011, S6-S7).
- unspecified: disable ignores rawValue; stored array bits may remain but count defines validity.
*)

IF enable THEN
    IF tmp_count < 8 THEN
        tmp_buffer[tmp_count] := rawValue;
        tmp_count := tmp_count + 1;
        IF tmp_count < 8 THEN
            tmp_write_index := tmp_count;
        ELSE
            tmp_write_index := 0;
        END_IF;
    ELSE
        tmp_buffer[tmp_write_index] := rawValue;
        tmp_write_index := tmp_write_index + 1;
        IF tmp_write_index > 7 THEN
            tmp_write_index := 0;
        END_IF;
    END_IF;

    tmp_sum := 0.0;
    FOR tmp_i := 0 TO tmp_count - 1 DO
        tmp_sum := tmp_sum + tmp_buffer[tmp_i];
    END_FOR;

    IF tmp_count > 0 THEN
        filteredValue := tmp_sum / INT_TO_REAL(tmp_count);
    END_IF;

    sampleCount := tmp_count;
    windowFull := (tmp_count = 8);
ELSE
    tmp_count := 0;
    tmp_write_index := 0;
    sampleCount := 0;
    windowFull := FALSE;
END_IF;

(* CONTRACT_RULES [] *)

END_FUNCTION_BLOCK

(* ---- self-medium-03.candidate_01.st ---- *)
(*
ENGINEERING_CONTRACT
- motorUp: start on IDLE open-button rising edge with closeBtn FALSE and openLimit FALSE; retain while moving; stop on obstacle/openLimit/fault/clear scan.
- motorDown: symmetric with openBtn FALSE and closeLimit FALSE; mutually exclusive with motorUp.
- errorFlag: set by any obstacle; latched; cleared only by no-obstacle rising(openBtn AND closeBtn); clear scan keeps motors off.
- State: initial IDLE; OPENING/CLOSING track active motion; FAULT latches; clear returns IDLE. Conflicting dual-button edge starts neither motor.
- Same-scan priority: obstacle/fault dominates limit, motion, and reset; outputs are evaluated from the current sampled inputs.
*)
(* CONTRACT_RULES [] *)

TYPE FB_STATE : (IDLE, OPENING, CLOSING, FAULT); END_TYPE;

FUNCTION_BLOCK FB
VAR_INPUT
    openBtn : BOOL;
    closeBtn : BOOL;
    openLimit : BOOL;
    closeLimit : BOOL;
    obstacle : BOOL;
END_VAR
VAR_OUTPUT
    motorUp : BOOL;
    motorDown : BOOL;
    errorFlag : BOOL;
END_VAR
VAR
    state : FB_STATE := FB_STATE#IDLE;
    prevOpenBtn : BOOL := FALSE;
    prevCloseBtn : BOOL := FALSE;
    prevMotorUp : BOOL := FALSE;
    prevMotorDown : BOOL := FALSE;
    prevErrorFlag : BOOL := FALSE;
    local_risingOpen : BOOL := FALSE;
    local_risingClose : BOOL := FALSE;
    local_risingBoth : BOOL := FALSE;
    local_errNow : BOOL := FALSE;
    local_startUp : BOOL := FALSE;
    local_startDown : BOOL := FALSE;
    local_runUp : BOOL := FALSE;
    local_runDown : BOOL := FALSE;
END_VAR

local_risingOpen := openBtn AND NOT prevOpenBtn;
local_risingClose := closeBtn AND NOT prevCloseBtn;
local_risingBoth := openBtn AND closeBtn AND NOT (prevOpenBtn AND prevCloseBtn);

local_errNow := obstacle OR (prevErrorFlag AND NOT local_risingBoth);

IF local_errNow THEN
    errorFlag := TRUE;
    motorUp := FALSE;
    motorDown := FALSE;
    state := FB_STATE#FAULT;
ELSE
    local_startUp := NOT prevMotorUp AND NOT prevMotorDown AND NOT prevErrorFlag
        AND NOT obstacle AND local_risingOpen AND NOT closeBtn AND NOT openLimit;
    local_startDown := NOT prevMotorUp AND NOT prevMotorDown AND NOT prevErrorFlag
        AND NOT obstacle AND local_risingClose AND NOT openBtn AND NOT closeLimit;
    local_runUp := prevMotorUp AND NOT prevErrorFlag AND NOT obstacle AND NOT openLimit;
    local_runDown := prevMotorDown AND NOT prevErrorFlag AND NOT obstacle AND NOT closeLimit;

    motorUp := local_startUp OR local_runUp;
    motorDown := local_startDown OR local_runDown;
    errorFlag := FALSE;

    IF motorUp THEN
        state := FB_STATE#OPENING;
    ELSIF motorDown THEN
        state := FB_STATE#CLOSING;
    ELSE
        state := FB_STATE#IDLE;
    END_IF;
END_IF;

prevOpenBtn := openBtn;
prevCloseBtn := closeBtn;
prevMotorUp := motorUp;
prevMotorDown := motorDown;
prevErrorFlag := errorFlag;

END_FUNCTION_BLOCK

(* ---- self-medium-03.candidate_03.st ---- *)
(*
ENGINEERING_CONTRACT
- motorUp: start on IDLE open-button rising edge with closeBtn FALSE and openLimit FALSE; retain while moving; stop on obstacle/openLimit/fault/clear scan.
- motorDown: symmetric with openBtn FALSE and closeLimit FALSE; mutually exclusive with motorUp.
- errorFlag: set by any obstacle; latched; cleared only by no-obstacle rising(openBtn AND closeBtn); clear scan keeps motors off.
- State: initial IDLE; OPENING/CLOSING track active motion; FAULT latches; clear returns IDLE. Conflicting dual-button edge starts neither motor.
- Same-scan priority: obstacle/fault dominates limit, motion, and reset; outputs are evaluated from the current sampled inputs.
*)
(* CONTRACT_RULES [] *)

TYPE FB_STATE : (IDLE, OPENING, CLOSING, FAULT); END_TYPE;

FUNCTION_BLOCK FB
VAR_INPUT
    openBtn : BOOL;
    closeBtn : BOOL;
    openLimit : BOOL;
    closeLimit : BOOL;
    obstacle : BOOL;
END_VAR
VAR_OUTPUT
    motorUp : BOOL;
    motorDown : BOOL;
    errorFlag : BOOL;
END_VAR
VAR
    state : FB_STATE := IDLE;
    prevOpenBtn : BOOL := FALSE;
    prevCloseBtn : BOOL := FALSE;
    prevMotorUp : BOOL := FALSE;
    prevMotorDown : BOOL := FALSE;
    prevErrorFlag : BOOL := FALSE;
    local_risingOpen : BOOL := FALSE;
    local_risingClose : BOOL := FALSE;
    local_risingBoth : BOOL := FALSE;
    local_errNow : BOOL := FALSE;
    local_startUp : BOOL := FALSE;
    local_startDown : BOOL := FALSE;
    local_runUp : BOOL := FALSE;
    local_runDown : BOOL := FALSE;
END_VAR

local_risingOpen := openBtn AND NOT prevOpenBtn;
local_risingClose := closeBtn AND NOT prevCloseBtn;
local_risingBoth := openBtn AND closeBtn AND NOT (prevOpenBtn AND prevCloseBtn);

local_errNow := obstacle OR (prevErrorFlag AND NOT local_risingBoth);

IF local_errNow THEN
    errorFlag := TRUE;
    motorUp := FALSE;
    motorDown := FALSE;
    state := FAULT;
ELSE
    local_startUp := NOT prevMotorUp AND NOT prevMotorDown AND NOT prevErrorFlag
        AND NOT obstacle AND local_risingOpen AND NOT closeBtn AND NOT openLimit;
    local_startDown := NOT prevMotorUp AND NOT prevMotorDown AND NOT prevErrorFlag
        AND NOT obstacle AND local_risingClose AND NOT openBtn AND NOT closeLimit;
    local_runUp := prevMotorUp AND NOT prevErrorFlag AND NOT obstacle AND NOT openLimit;
    local_runDown := prevMotorDown AND NOT prevErrorFlag AND NOT obstacle AND NOT closeLimit;

    motorUp := local_startUp OR local_runUp;
    motorDown := local_startDown OR local_runDown;
    errorFlag := FALSE;

    IF motorUp THEN
        state := OPENING;
    ELSIF motorDown THEN
        state := CLOSING;
    ELSE
        state := IDLE;
    END_IF;
END_IF;

prevOpenBtn := openBtn;
prevCloseBtn := closeBtn;
prevMotorUp := motorUp;
prevMotorDown := motorDown;
prevErrorFlag := errorFlag;

END_FUNCTION_BLOCK

(* ---- self-medium-03.patch_base_03.st ---- *)
(*
ENGINEERING_CONTRACT
- motorUp: start on IDLE open-button rising edge with closeBtn FALSE and openLimit FALSE; retain while moving; stop on obstacle/openLimit/fault/clear scan.
- motorDown: symmetric with openBtn FALSE and closeLimit FALSE; mutually exclusive with motorUp.
- errorFlag: set by any obstacle; latched; cleared only by no-obstacle rising(openBtn AND closeBtn); clear scan keeps motors off.
- State: initial IDLE; OPENING/CLOSING track active motion; FAULT latches; clear returns IDLE. Conflicting dual-button edge starts neither motor.
- Same-scan priority: obstacle/fault dominates limit, motion, and reset; outputs are evaluated from the current sampled inputs.
*)
(* CONTRACT_RULES [] *)

TYPE FB_STATE : (IDLE, OPENING, CLOSING, FAULT); END_TYPE;

FUNCTION_BLOCK FB
VAR_INPUT
    openBtn : BOOL;
    closeBtn : BOOL;
    openLimit : BOOL;
    closeLimit : BOOL;
    obstacle : BOOL;
END_VAR
VAR_OUTPUT
    motorUp : BOOL;
    motorDown : BOOL;
    errorFlag : BOOL;
END_VAR
VAR
    state : FB_STATE := FB_STATE#IDLE;
    prevOpenBtn : BOOL := FALSE;
    prevCloseBtn : BOOL := FALSE;
    prevMotorUp : BOOL := FALSE;
    prevMotorDown : BOOL := FALSE;
    prevErrorFlag : BOOL := FALSE;
    local_risingOpen : BOOL := FALSE;
    local_risingClose : BOOL := FALSE;
    local_risingBoth : BOOL := FALSE;
    local_errNow : BOOL := FALSE;
    local_startUp : BOOL := FALSE;
    local_startDown : BOOL := FALSE;
    local_runUp : BOOL := FALSE;
    local_runDown : BOOL := FALSE;
END_VAR

local_risingOpen := openBtn AND NOT prevOpenBtn;
local_risingClose := closeBtn AND NOT prevCloseBtn;
local_risingBoth := openBtn AND closeBtn AND NOT (prevOpenBtn AND prevCloseBtn);

local_errNow := obstacle OR (prevErrorFlag AND NOT local_risingBoth);

IF local_errNow THEN
    errorFlag := TRUE;
    motorUp := FALSE;
    motorDown := FALSE;
    state := FB_STATE#FAULT;
ELSE
    local_startUp := NOT prevMotorUp AND NOT prevMotorDown AND NOT prevErrorFlag
        AND NOT obstacle AND local_risingOpen AND NOT closeBtn AND NOT openLimit;
    local_startDown := NOT prevMotorUp AND NOT prevMotorDown AND NOT prevErrorFlag
        AND NOT obstacle AND local_risingClose AND NOT openBtn AND NOT closeLimit;
    local_runUp := prevMotorUp AND NOT prevErrorFlag AND NOT obstacle AND NOT openLimit;
    local_runDown := prevMotorDown AND NOT prevErrorFlag AND NOT obstacle AND NOT closeLimit;

    motorUp := local_startUp OR local_runUp;
    motorDown := local_startDown OR local_runDown;
    errorFlag := FALSE;

    IF motorUp THEN
        state := FB_STATE#OPENING;
    ELSIF motorDown THEN
        state := FB_STATE#CLOSING;
    ELSE
        state := FB_STATE#IDLE;
    END_IF;
END_IF;

prevOpenBtn := openBtn;
prevCloseBtn := closeBtn;
prevMotorUp := motorUp;
prevMotorDown := motorDown;
prevErrorFlag := errorFlag;

END_FUNCTION_BLOCK

(* ---- self-medium-03.raw_candidate_01.st ---- *)
(*
ENGINEERING_CONTRACT
- motorUp: start on IDLE open-button rising edge with closeBtn FALSE and openLimit FALSE; retain while moving; stop on obstacle/openLimit/fault/clear scan.
- motorDown: symmetric with openBtn FALSE and closeLimit FALSE; mutually exclusive with motorUp.
- errorFlag: set by any obstacle; latched; cleared only by no-obstacle rising(openBtn AND closeBtn); clear scan keeps motors off.
- State: initial IDLE; OPENING/CLOSING track active motion; FAULT latches; clear returns IDLE. Conflicting dual-button edge starts neither motor.
- Same-scan priority: obstacle/fault dominates limit, motion, and reset; outputs are evaluated from the current sampled inputs.
*)
(* CONTRACT_RULES [] *)

TYPE FB_STATE : (IDLE, OPENING, CLOSING, FAULT); END_TYPE

FUNCTION_BLOCK FB
VAR_INPUT
    openBtn : BOOL;
    closeBtn : BOOL;
    openLimit : BOOL;
    closeLimit : BOOL;
    obstacle : BOOL;
END_VAR
VAR_OUTPUT
    motorUp : BOOL;
    motorDown : BOOL;
    errorFlag : BOOL;
END_VAR
VAR
    state : FB_STATE := FB_STATE#IDLE;
    prevOpenBtn : BOOL := FALSE;
    prevCloseBtn : BOOL := FALSE;
    prevMotorUp : BOOL := FALSE;
    prevMotorDown : BOOL := FALSE;
    prevErrorFlag : BOOL := FALSE;
    local_risingOpen : BOOL := FALSE;
    local_risingClose : BOOL := FALSE;
    local_risingBoth : BOOL := FALSE;
    local_errNow : BOOL := FALSE;
    local_startUp : BOOL := FALSE;
    local_startDown : BOOL := FALSE;
    local_runUp : BOOL := FALSE;
    local_runDown : BOOL := FALSE;
END_VAR

local_risingOpen := openBtn AND NOT prevOpenBtn;
local_risingClose := closeBtn AND NOT prevCloseBtn;
local_risingBoth := openBtn AND closeBtn AND NOT (prevOpenBtn AND prevCloseBtn);

local_errNow := obstacle OR (prevErrorFlag AND NOT local_risingBoth);

IF local_errNow THEN
    errorFlag := TRUE;
    motorUp := FALSE;
    motorDown := FALSE;
    state := FB_STATE#FAULT;
ELSE
    local_startUp := NOT prevMotorUp AND NOT prevMotorDown AND NOT prevErrorFlag
        AND NOT obstacle AND local_risingOpen AND NOT closeBtn AND NOT openLimit;
    local_startDown := NOT prevMotorUp AND NOT prevMotorDown AND NOT prevErrorFlag
        AND NOT obstacle AND local_risingClose AND NOT openBtn AND NOT closeLimit;
    local_runUp := prevMotorUp AND NOT prevErrorFlag AND NOT obstacle AND NOT openLimit;
    local_runDown := prevMotorDown AND NOT prevErrorFlag AND NOT obstacle AND NOT closeLimit;

    motorUp := local_startUp OR local_runUp;
    motorDown := local_startDown OR local_runDown;
    errorFlag := FALSE;

    IF motorUp THEN
        state := FB_STATE#OPENING;
    ELSIF motorDown THEN
        state := FB_STATE#CLOSING;
    ELSE
        state := FB_STATE#IDLE;
    END_IF;
END_IF;

prevOpenBtn := openBtn;
prevCloseBtn := closeBtn;
prevMotorUp := motorUp;
prevMotorDown := motorDown;
prevErrorFlag := errorFlag;

END_FUNCTION_BLOCK

(* ---- self-medium-03.raw_candidate_03.st ---- *)
(*
ENGINEERING_CONTRACT
- motorUp: start on IDLE open-button rising edge with closeBtn FALSE and openLimit FALSE; retain while moving; stop on obstacle/openLimit/fault/clear scan.
- motorDown: symmetric with openBtn FALSE and closeLimit FALSE; mutually exclusive with motorUp.
- errorFlag: set by any obstacle; latched; cleared only by no-obstacle rising(openBtn AND closeBtn); clear scan keeps motors off.
- State: initial IDLE; OPENING/CLOSING track active motion; FAULT latches; clear returns IDLE. Conflicting dual-button edge starts neither motor.
- Same-scan priority: obstacle/fault dominates limit, motion, and reset; outputs are evaluated from the current sampled inputs.
*)
(* CONTRACT_RULES [] *)

TYPE FB_STATE : (IDLE, OPENING, CLOSING, FAULT); END_TYPE;

FUNCTION_BLOCK FB
VAR_INPUT
    openBtn : BOOL;
    closeBtn : BOOL;
    openLimit : BOOL;
    closeLimit : BOOL;
    obstacle : BOOL;
END_VAR
VAR_OUTPUT
    motorUp : BOOL;
    motorDown : BOOL;
    errorFlag : BOOL;
END_VAR
VAR
    state : FB_STATE := IDLE;
    prevOpenBtn : BOOL := FALSE;
    prevCloseBtn : BOOL := FALSE;
    prevMotorUp : BOOL := FALSE;
    prevMotorDown : BOOL := FALSE;
    prevErrorFlag : BOOL := FALSE;
    local_risingOpen : BOOL := FALSE;
    local_risingClose : BOOL := FALSE;
    local_risingBoth : BOOL := FALSE;
    local_errNow : BOOL := FALSE;
    local_startUp : BOOL := FALSE;
    local_startDown : BOOL := FALSE;
    local_runUp : BOOL := FALSE;
    local_runDown : BOOL := FALSE;
END_VAR

local_risingOpen := openBtn AND NOT prevOpenBtn;
local_risingClose := closeBtn AND NOT prevCloseBtn;
local_risingBoth := openBtn AND closeBtn AND NOT (prevOpenBtn AND prevCloseBtn);

local_errNow := obstacle OR (prevErrorFlag AND NOT local_risingBoth);

IF local_errNow THEN
    errorFlag := TRUE;
    motorUp := FALSE;
    motorDown := FALSE;
    state := FAULT;
ELSE
    local_startUp := NOT prevMotorUp AND NOT prevMotorDown AND NOT prevErrorFlag
        AND NOT obstacle AND local_risingOpen AND NOT closeBtn AND NOT openLimit;
    local_startDown := NOT prevMotorUp AND NOT prevMotorDown AND NOT prevErrorFlag
        AND NOT obstacle AND local_risingClose AND NOT openBtn AND NOT closeLimit;
    local_runUp := prevMotorUp AND NOT prevErrorFlag AND NOT obstacle AND NOT openLimit;
    local_runDown := prevMotorDown AND NOT prevErrorFlag AND NOT obstacle AND NOT closeLimit;

    motorUp := local_startUp OR local_runUp;
    motorDown := local_startDown OR local_runDown;
    errorFlag := FALSE;

    IF motorUp THEN
        state := OPENING;
    ELSIF motorDown THEN
        state := CLOSING;
    ELSE
        state := IDLE;
    END_IF;
END_IF;

prevOpenBtn := openBtn;
prevCloseBtn := closeBtn;
prevMotorUp := motorUp;
prevMotorDown := motorDown;
prevErrorFlag := errorFlag;

END_FUNCTION_BLOCK

(* ---- self-medium-04.candidate_01.st ---- *)
FUNCTION_BLOCK FB
VAR_INPUT
    startBtn   : BOOL;
    resetBtn   : BOOL;
    doneSensor : BOOL;
    targetVol  : REAL;
    flowVol    : REAL;
END_VAR
VAR_OUTPUT
    valveOpen  : BOOL;
    fillsToday : INT;
END_VAR
VAR
    prevStartBtn   : BOOL := FALSE;
    prevResetBtn   : BOOL := FALSE;
    prevValveOpen  : BOOL := FALSE;
    pendingConfirm : BOOL := FALSE;
    accumulatedVol : REAL := 0.0;
    tmp_risingReset : BOOL;
    tmp_risingStart : BOOL;
    tmp_isFilling   : BOOL;
END_VAR

(* ENGINEERING_CONTRACT
   valveOpen: set only on start edge from idle/wait (R2,S2); holds while
             accumulatedVol < targetVol (R3,S9); closes on reset or target reach (R1,R3,S5).
   pendingConfirm: set same scan as target close; persists until confirmation,
             next start, or reset; sensor TRUE does not repeat count (R3-R5,S11).
   fillsToday: increments once on doneSensor with pending; saturates at 32767
             and still clears pending; reset zeros in same scan (R4-R5,S1,S6,S14).
   accumulatedVol: reset on reset/new bottle; adds flowVol only while filling,
             including start scan (R1-R3,S12).
   Priority: reset > start/new-bottle cancellation > flow/threshold close > done confirm.
   Units: targetVol/flowVol in mL REAL; fillsToday signed INT bounds 0..32767.
*)

(* CONTRACT_RULES [] *)

tmp_risingReset := resetBtn AND NOT prevResetBtn;
tmp_risingStart := startBtn AND NOT prevStartBtn;

IF tmp_risingReset THEN
    valveOpen      := FALSE;
    fillsToday     := 0;
    accumulatedVol := 0.0;
    pendingConfirm := FALSE;
ELSE
    tmp_isFilling := FALSE;

    IF tmp_risingStart AND NOT valveOpen THEN
        pendingConfirm := FALSE;
        accumulatedVol := 0.0;
        valveOpen      := TRUE;
        tmp_isFilling   := TRUE;
    ELSIF valveOpen THEN
        tmp_isFilling := TRUE;
    END_IF;

    IF tmp_isFilling THEN
        accumulatedVol := accumulatedVol + flowVol;
        IF accumulatedVol >= targetVol THEN
            valveOpen      := FALSE;
            pendingConfirm := TRUE;
            tmp_isFilling   := FALSE;
        END_IF;
    END_IF;

    IF pendingConfirm AND doneSensor THEN
        IF fillsToday < 32767 THEN
            fillsToday := fillsToday + 1;
        END_IF;
        pendingConfirm := FALSE;
    END_IF;
END_IF;

prevStartBtn  := startBtn;
prevResetBtn  := resetBtn;
prevValveOpen := valveOpen;

END_FUNCTION_BLOCK
